(* IEC 61131-3 sources: daoli-st-library/DL_Device (part 35) *)

(* ---- FB_DL_ValveSeatLeakWatch.st ---- *)
(*==============================================================================
 * 组件名称 (Component)  : FB_DL_ValveSeatLeakWatch
 * 所属子库 (Sublibrary) : DL_Device
 * 当前版本 (Version)    : 1.0.1
 * 兼容性 (Platform)     : CODESYS 3.5+ / TwinCAT 3 / 汇川 InoProShop / 施耐德 Machine Expert
 *                         仅依赖 Standard.library（TON / R_TRIG），零厂商私有库
 * 功能描述 (Function)   : 阀座关闭位泄漏趋势监视。阀门命令关 + 关位反馈到齐 +
 *                         tSettle 稳定后进入监视：对关位残差（dp 或流量）做
 *                         N 点最小二乘趋势斜率（窗口线性回归）+ 均值双判据：
 *                         残差均值超 fLeakLevel 且斜率非负上升 → 泄漏判据成立，
 *                         bLeakDetected 锁存。开阀/离开关位自动回监视待机。
 * 来源标签 (Origin)     : 自研线（诊断族深化，IEC 61131-3 标准语义的道莅防御性
 *                         实现，clean-room）
 * 分工声明 (Pairing)    : ValveSeatLeakWatch（关位泄漏趋势，本件）↔
 *                         ValvePartialStrokeTest（行程试验，既有件）：本件只在
 *                         关位做无扰动趋势监视，不驱动阀门动作；行程试验主动
 *                         部分行程激励，二者判据域不同不互斥（R298 属主边界）。
 * 边界语义 (Boundary)   : ① 判据串相位因子：仅 eWatch 相判泄漏，eIdle/开阀期
 *                         不判（R281 相位相关判据防误锁口径）；
 *                         ② LS 除零防御：Σ(x-x̄)² <= eps（窗口内无时间跨度）
 *                         → 斜率按 0 处理，只走均值判据，不产生 Inf；
 *                         ③ 残差 NaN 拒收（不入窗口，不参与统计）；
 *                         ④ 组态闸：窗深 < 2 / 阈值 <= 0 / 稳定时间 <= 0 → 故障。
 * 输出语义 (Fallback)   : 【R191】eIdle 相 → 判据输出清零（监视未在关位，
 *                         无泄漏语义）；eFault 相 → bLeakDetected 保持末值 +
 *                         bError = TRUE。
 * 码位     (Codes)      : 按 R297 范式零 16# 码位硬编码；错误出口 BOOL+ENUM(eCause)，
 *                         码位待主控收口统一派号。
 * 红线自检 (Redline)    : 7 项红线已自检：R1 零全局 ✓｜R2 零物理地址 ✓｜R3 纯 IEC ✓
 *                         R4 除零（Σx² eps 闸）/NaN 拒收/组态闸 ✓
 *                         R5 双语同行注释 ✓｜R6 CASE 带 ELSE 兜底迁 eFault ✓
 *                         R7 TON/R_TRIG 段 0 无条件刷新，各自独立实例 ✓
 * 验收向量 (Acceptance) : V1 关位稳定后残差恒 0.5（阈 0.2）、窗口斜率 ≈ 0 →
 *                         斜率非负成立，tLeakConf 到时 bLeakDetected=TRUE；
 *                         V2 残差 0.5 但窗口斜率显著负下降 → 不判泄漏；
 *                         V3 开阀命令一出现 → 判据清零回 eIdle。
 * 修订历史 (Revision)   : 2026-11-20  v1.0.0  R49 首版（批 2 · 序号 8）
 *                        2026-11-20  v1.0.1  R52: 环窗时间序修正，消除斜率符号翻转
 *                        （删写入期 _aX[_nHead] 赋值，改求和期按 _nOldest→_nIdx 时间序
 *                        环回取 _aRes，X 用 1.._nFill 时间序号；修回卷后 X/Y 错配致
 *                        L193 `_fSlope >= 0.0` 把真实上升泄漏判成非上升的安全侧漏报）
 *==============================================================================*)
TYPE E_DL_VslState :
(
    eIdle   := 0,                            (* 未在关位（判据清零） / Not at closed seat *)
    eSettle := 10,                           (* 关位稳定等待 / Closed-seat settling *)
    eWatch  := 20,                           (* 泄漏趋势监视 / Leak trend watching *)
    eFault  := 90                            (* 故障锁存相 / Fault latched phase *)
);
END_TYPE

TYPE E_DL_VslCause :
(
    eNone       := 0,                        (* 无故障成因 / No cause *)
    eCfgIllegal := 1,                        (* 组态非法：窗深/阈值/时间越域 / Illegal config *)
    ePhaseBad   := 2                         (* 非法相位兜底 / Illegal phase fallback *)
);
END_TYPE

FUNCTION_BLOCK FB_DL_ValveSeatLeakWatch
VAR_INPUT
    bCmdClose   : BOOL := FALSE;             (* 阀关命令电平 [-] / Valve close command level *)
    bLimitClosed: BOOL := FALSE;             (* 关位限位反馈电平 [-] / Closed-seat limit feedback *)
    fResidual   : LREAL := 0.0;              (* 关位残差输入（dp 或流量标定值）[工程单位] / Closed-seat residual input *)
    fLeakLevel  : LREAL := 0.2;              (* 泄漏均值阈值，域 > 0.0 [工程单位] / Leak mean threshold *)
    nWinDepth   : INT := 16;                 (* LS 趋势窗深，域 2..32 [点] / LS trend window depth *)
    tSettle     : TIME := T#5S;              (* 关位稳定等待时间，域 > T#0S [ms] / Settle wait time *)
    tLeakConf   : TIME := T#3S;              (* 泄漏判据确认保持时间，域 > T#0S [ms] / Leak confirm hold time *)
    bEnable     : BOOL := TRUE;              (* 监视使能 [-] / Enable *)
    bReset      : BOOL := FALSE;             (* 复位命令，上升沿清泄漏锁存与窗口 [-] / Reset command *)
END_VAR
VAR_OUTPUT
    bLeakDetected : BOOL;                    (* 泄漏判据锁存位（复位沿或开阀沿清）[-] / Leak detected latch *)
    fResidualMean : LREAL;                   (* 当前窗口残差均值 [工程单位] / Window residual mean *)
    fTrendSlope   : LREAL;                   (* 当前窗口 LS 趋势斜率 [工程单位/拍] / Window LS slope *)
    bWatching     : BOOL;                    (* 关位监视中指示 [-] / Watching indicator *)
    eState        : E_DL_VslState;           (* 状态出口 / State outlet *)
    eCause        : E_DL_VslCause;           (* 故障成因出口（R190 归因唯一） / Fault cause outlet *)
    bError        : BOOL;                    (* 故障锁存标志 [-] / Fault latch flag *)
END_VAR
VAR
    _eState  : E_DL_VslState := E_DL_VslState.eIdle;      (* 内部相位（CASE 唯一写入目标） / Internal phase *)
    _eCause  : E_DL_VslCause := E_DL_VslCause.eNone;      (* 故障成因锁存量 / Latched cause *)
    tonSettle: TON;                          (* 关位稳定计时，IN 由相位派生，段 0 无条件调用 / Settle timer *)
    tonConf  : TON;                          (* 泄漏确认计时，独立实例（一相一定时器，R275） / Confirm timer, separate instance *)
    rtReset  : R_TRIG;                       (* 复位沿实例，段 0 无条件调用 / Reset edge instance *)
    _aRes    : ARRAY[1..32] OF LREAL;        (* 残差窗口环形缓冲 [工程单位] / Residual ring window *)
    _aX      : ARRAY[1..32] OF LREAL;        (* 窗口序号数组（v1.0.1 起废弃不参与运算，R53 清理；保留以保差异审阅可读）[点] / Deprecated index array *)
    _nHead   : INT;                          (* 环形写入头游标 [-] / Ring head cursor *)
    _nOldest : INT;                          (* 最旧样本槽位（统计段每趟重算）[-] / Oldest sample slot, recomputed *)
    _nIdx    : INT;                          (* 时间序 → 环形槽位换算下标 [-] / Time-order to slot index *)
    _nFill   : INT;                          (* 窗口已填充点数 [点] / Window fill count *)
    _nEff    : INT;                          (* 钳位后生效窗深 [点] / Clamped effective depth *)
    _fSumX   : LREAL;                        (* LS 累计：Σx [-] / LS sum of x *)
    _fSumY   : LREAL;                        (* LS 累计：Σy [工程单位] / LS sum of y *)
    _fSumXY  : LREAL;                        (* LS 累计：Σxy [工程单位·点] / LS sum of xy *)
    _fSumX2  : LREAL;                        (* LS 累计：Σx² [-] / LS sum of x² *)
    _fDen    : LREAL;                        (* LS 分母 Σ(x-x̄)² [-] / LS denominator *)
    _fSlope  : LREAL;                        (* 本拍派生斜率 [工程单位/点] / Derived slope *)
    _fMean   : LREAL;                        (* 本拍派生均值 [工程单位] / Derived mean *)
    _bLeakC  : BOOL;                         (* 泄漏当拍判据（均值超阈 ∧ 斜率非负） / Leak verdict this scan *)
    _bFault  : BOOL;                         (* 故障锁存位 / Latched fault bit *)
    _bCfgBad : BOOL;                         (* 组态非法当拍量 / Illegal config this scan *)
    _i       : INT;                          (* 统计扫描游标（每趟重置，R227）[-] / Stats scan cursor *)
END_VAR
VAR CONSTANT
    DL_VSL_EPS  : LREAL := 1.0E-12;          (* LS 分母判零容差 [-] / LS denominator epsilon *)
    DL_VSL_NMAX : INT   := 32;               (* 窗深容量上限 [点] / Window capacity limit *)
END_VAR

(* —— 段 0：当拍判据派生 + 实例无条件刷新（R228A） —— *)
_bCfgBad := (fLeakLevel <= 0.0) OR (tSettle <= T#0S) OR (tLeakConf <= T#0S);   (* 组态闸（标量域引脚，R151） / Config gate *)
rtReset(CLK := bReset);                                                       (* 复位沿每拍必调 / Reset edge every scan *)
tonSettle(IN := _eState = E_DL_VslState.eSettle, PT := tSettle);              (* 稳定计时随相位派生 / Settle timer *)
tonConf(IN := _bLeakC AND _eState = E_DL_VslState.eWatch, PT := tLeakConf);   (* 确认计时（注意：IN 引用上拍判据，一拍滞后可接受，头注释声明） / Confirm timer, one-scan lag declared *)
_nEff := nWinDepth;                                                           (* 生效窗深初值 / Effective depth init *)
IF _nEff < 2 THEN
    _nEff := 2;                                                               (* 窗深下限 2（两点才能定斜率） / Min depth 2 *)
END_IF
IF _nEff > DL_VSL_NMAX THEN
    _nEff := DL_VSL_NMAX;                                                     (* 窗深钳位到容量（R308） / Clamp depth to capacity *)
END_IF
IF (nWinDepth < 2) OR (nWinDepth > DL_VSL_NMAX) THEN
    _bCfgBad := _bCfgBad OR TRUE;                                             (* 窗深越域并入组态闸（越域仍钳位运行但报故障） / Depth out of domain joins gate *)
END_IF

(* —— 段 1：单拍量预清零（R107） —— *)
_bLeakC := FALSE;                                                             (* 泄漏当拍判据预清，唯一分支置位 / Leak verdict preset *)
_fSumX := 0.0;                                                                (* LS 累计量清零重算（每拍全路径派生） / LS sums recompute *)
_fSumY := 0.0;                                                                (* Σy 清零 / Sum y clear *)
_fSumXY := 0.0;                                                               (* Σxy 清零 / Sum xy clear *)
_fSumX2 := 0.0;                                                               (* Σx² 清零 / Sum x2 clear *)
_fDen := 0.0;                                                                 (* LS 分母清零（防 _nFill=0 时旧值残留触发除零） / LS denominator clear *)
_fSlope := 0.0;                                                               (* 斜率缺省 0 / Slope default *)
_fMean := 0.0;                                                                (* 均值缺省 0 / Mean default *)
_nOldest := 1;                                                                (* 最旧槽位预清（统计段重算，防残留） / Oldest slot preset *)
_nIdx := 1;                                                                   (* 槽位下标预清 / Slot index preset *)

(* —— 段 2：复位沿处理（作用域：清故障 + 清泄漏锁存 + 清窗口 + 迁 eIdle，R283 逐项声明） —— *)
IF rtReset.Q THEN
    _bFault := FALSE;                                                         (* 清故障锁存 / Clear fault *)
    _eCause := E_DL_VslCause.eNone;                                           (* 清成因 / Clear cause *)
    bLeakDetected := FALSE;                                                   (* 清泄漏锁存 / Clear leak latch *)
    _nFill := 0;                                                              (* 清窗填充计数 / Clear fill count *)
    _nHead := 1;                                                              (* 头游标复位 / Head cursor reset *)
    _eState := E_DL_VslState.eIdle;                                           (* 迁待机相 / Back to idle *)
END_IF

(* —— 段 3：CASE 主状态机（判据串相位因子，R281；ELSE 兜底迁 eFault，红线 6） —— *)
CASE _eState OF
    E_DL_VslState.eIdle:                                                      (* 待机相：判据与统计出口清零（声明语义） / Idle: verdicts cleared *)
        fResidualMean := 0.0;                                                 (* 均值出口清零 / Mean outlet clear *)
        fTrendSlope := 0.0;                                                   (* 斜率出口清零 / Slope outlet clear *)
        bLeakDetected := FALSE;                                               (* 泄漏锁存随离开关位自动清（声明：开阀沿清锁存） / Leak latch auto-clear on leaving seat *)
        IF bEnable AND NOT _bFault AND bCmdClose AND bLimitClosed THEN
            _eState := E_DL_VslState.eSettle;                                 (* 关位到齐进入稳定等待 / Enter settle *)
        END_IF
    E_DL_VslState.eSettle:                                                    (* 稳定等待相 / Settle *)
        IF NOT (bCmdClose AND bLimitClosed) THEN
            _eState := E_DL_VslState.eIdle;                                   (* 离开关位回待机 / Leave seat *)
        ELSIF tonSettle.Q THEN
            _nFill := 0;                                                      (* 稳定后清窗重采（避免稳定前残差污染统计） / Clear window after settle *)
            _nHead := 1;                                                      (* 头游标复位 / Head reset *)
            _eState := E_DL_VslState.eWatch;                                  (* 进入监视 / Enter watch *)
        END_IF
    E_DL_VslState.eWatch:                                                     (* 监视相：采窗 + 统计 + 判据 / Watch *)
        IF NOT (bCmdClose AND bLimitClosed) THEN
            bLeakDetected := FALSE;                                           (* 离开位清泄漏锁存（开阀沿语义） / Leak latch clear *)
            _eState := E_DL_VslState.eIdle;                                   (* 回待机 / Back to idle *)
        ELSE
            IF (fResidual = fResidual) AND ((fResidual - fResidual) = (fResidual - fResidual)) THEN
                _aRes[_nHead] := fResidual;                                   (* 有限残差入环窗（NaN 拒收不入窗） / Finite residual into ring *)
                (* X 不再于写入期生成：改为求和期按时间序现算（R52 修 R193 扩面） / X derived at sum time in time order *)
                _nHead := _nHead + 1;                                         (* 头游标递进 / Head advance *)
                IF _nHead > _nEff THEN
                    _nHead := 1;                                              (* 环回卷（下标先判后增，无越界） / Ring wrap *)
                END_IF
                IF _nFill < _nEff THEN
                    _nFill := _nFill + 1;                                     (* 填充计数封顶 / Fill count cap *)
                END_IF
            END_IF
            IF _nFill >= 1 THEN
                _nOldest := _nHead - _nFill;                                  (* 最旧样本槽：未满窗时 = 1（头游标 = 填充数 + 1） / Oldest slot while filling *)
                IF _nOldest < 1 THEN
                    _nOldest := _nOldest + _nEff;                             (* 满窗回卷后最旧样本在 _nHead 槽：时间序起点（R52 修） / Wrapped: oldest at head slot *)
                END_IF
            END_IF
            _i := 1;                                                          (* 统计游标起头重置（R227） / Stats cursor reset *)
            WHILE _i <= _nFill DO                                             (* 逐点 LS 累计：x = 时间序，y 自最旧槽环回取值（R52 时间序） / Time-ordered LS sums *)
                _nIdx := _nOldest + _i - 1;                                   (* 时间序 → 环形槽位映射 / Time order to ring slot *)
                IF _nIdx > _nEff THEN
                    _nIdx := _nIdx - _nEff;                                   (* 槽位环回 / Slot wrap *)
                END_IF
                _fSumX := _fSumX + DINT_TO_LREAL(_i);                         (* Σx（时间序号 1..nFill，不随运行时间增长） / Sum x in time order *)
                _fSumY := _fSumY + _aRes[_nIdx];                              (* Σy / Sum y *)
                _fSumXY := _fSumXY + DINT_TO_LREAL(_i) * _aRes[_nIdx];        (* Σxy / Sum xy *)
                _fSumX2 := _fSumX2 + DINT_TO_LREAL(_i) * DINT_TO_LREAL(_i);   (* Σx² / Sum x2 *)
                _i := _i + 1;                                                 (* 游标递进 / Cursor advance *)
            END_WHILE
            IF _nFill >= 1 THEN
                _fMean := _fSumY / DINT_TO_LREAL(_nFill);                     (* 均值：除子恒 >= 1 无除零 / Mean, divisor >= 1 *)
                _fDen := _fSumX2 - _fSumX * _fSumX / DINT_TO_LREAL(_nFill);   (* LS 分母 = Σx² - (Σx)²/n / LS denominator *)
            END_IF
            IF _fDen > DL_VSL_EPS THEN
                _fSlope := (_fSumXY - _fSumX * _fSumY / DINT_TO_LREAL(_nFill)) / _fDen;   (* 斜率：分母已过 eps 闸，无除零 / Slope, denominator gated *)
            ELSE
                _fSlope := 0.0;                                               (* 窗内无时间跨度：斜率退化 0，只走均值判据（边界②） / Degenerate slope zero *)
            END_IF
            fResidualMean := _fMean;                                          (* 均值出口镜像 / Mean outlet mirror *)
            fTrendSlope := _fSlope;                                           (* 斜率出口镜像 / Slope outlet mirror *)
            _bLeakC := (_fMean > fLeakLevel) AND (_fSlope >= 0.0);            (* 判据：均值超阈 ∧ 斜率非负（0.0 容差比较：斜率与 0 用 >= 单侧合法） / Verdict: mean over threshold AND slope non-negative *)
            IF tonConf.Q THEN                                                 (* 判据保持到确认时间 / Verdict held to confirm time *)
                bLeakDetected := TRUE;                                        (* 泄漏锁存至复位沿/离开位 / Leak latch *)
            END_IF
        END_IF
    E_DL_VslState.eFault:                                                     (* 故障相：保持末值，仅复位沿出 / Fault *)
        ;                                                                     (* 锁存回放（R28） / Replay from latch *)
    ELSE                                                                      (* 非法相位兜底迁安全态 / Illegal phase fallback *)
        _eState := E_DL_VslState.eFault;                                      (* 迁故障相 / To fault *)
        _bFault := TRUE;                                                      (* 同步锁存 / Latch *)
        _eCause := E_DL_VslCause.ePhaseBad;                                   (* 成因：非法相位 / Cause: illegal phase *)
END_CASE

(* —— 段 4：出口映射（bError/eState 同源，R191） —— *)
bWatching := (_eState = E_DL_VslState.eWatch);                                (* 监视中指示 / Watching indicator *)
bError := _bFault;                                                            (* 故障标志镜像 / Fault flag mirror *)
eState := _eState;                                                            (* 状态出口 / State outlet *)
eCause := _eCause;                                                            (* 成因出口 / Cause outlet *)
END_FUNCTION_BLOCK

(* ---- FB_DL_ValveStrokeTimeWatch.st ---- *)
// FB_DL_ValveStrokeTimeWatch v1.0.0
(*==============================================================================
 * 功能描述: 阀门行程时间监视。开/关指令上升沿起 TON 计测，到限位反馈即记录
 *           本次行程时间 fStrokeTime [s]；行程未在 tMax 内到位 → bSlow 告警锁存；
 *           指令撤销（中途回退）即复位计时。开/关双向独立监视，bSlow 仅由 bReset
 *           复位沿解除（正常行程不清除既有告警）。
 * 接口契约: 输入 bOpenCmd/bCloseCmd/bOpenedLim/bClosedLim/tMax/bReset；
 *           输出 fStrokeTime/bSlow/bMoving/bError（恒假兼容出口）/nErrId。
 * 边界: ① 四枚 R_TRIG + 两枚 TON 段 0 无条件周期刷新；② 开/关命令互斥（同拍双真
 *           以开优先，暂不报专用码位）；③ tMax <= T#0S → 视为无效组态，PT 即时到
 *           时（bSlow 直告），恢复监视需改回有效组态；
 *           ④ 零全局耦合。
 * 码表: 16#0007_0309 信息级：慢行程告警（bSlow 并行，每拍重算）；故障相无锁存
 *       （bSlow 为告警级，随正常行程或复位沿解除）。
 * 修订历史: 2026-11-23  v1.0.0  R74 首版
 *==============================================================================*)

FUNCTION_BLOCK FB_DL_ValveStrokeTimeWatch
VAR_INPUT
    bOpenCmd   : BOOL := FALSE;    // 开阀指令 [-] / Open command
    bCloseCmd  : BOOL := FALSE;    // 关阀指令 [-] / Close command
    bOpenedLim : BOOL := FALSE;    // 开到位限位反馈 [-] / Opened limit feedback
    bClosedLim : BOOL := FALSE;    // 关到位限位反馈 [-] / Closed limit feedback
    tMax       : TIME := T#30S;    // 行程时间上限，域 > T#0S [ms] / Stroke time upper limit
    bReset     : BOOL := FALSE;    // 复位，上升沿清 bSlow 锁存 [-] / Reset edge clears slow latch
END_VAR
VAR_OUTPUT
    fStrokeTime : REAL := 0.0;     // 最近一次完成行程时间 [s] / Last completed stroke time [s]
    bSlow       : BOOL;            // 慢行程告警锁存 [-] / Slow stroke latch
    bMoving     : BOOL;            // 行进中标志（指令且未到限位）[-] / Moving flag
    bError      : BOOL;            // 故障锁存出口（本件无故障级，恒假，兼容出口口径）[-] / Fault outlet, always FALSE here
    nErrId      : UDINT;           // 事件码，0 = 无事件 / Event code, 0 = none
END_VAR
VAR
    rtOpen    : R_TRIG;            // 开指令上升沿实例，段 0 无条件刷新 / Open command rising edge
    rtClose   : R_TRIG;            // 关指令上升沿实例，段 0 无条件刷新 / Close command rising edge
    rtReset   : R_TRIG;            // 复位沿实例，段 0 无条件刷新 / Reset edge instance
    tonOpen   : TON;               // 开行程计时，段 0 无条件刷新 / Open stroke timer
    tonClose  : TON;               // 关行程计时，段 0 无条件刷新 / Close stroke timer
    _bCfgBad  : BOOL;              // 组态非法当拍量 [-] / Illegal configuration this scan
    _bCmdDual : BOOL;              // 开关命令同拍双真当拍量 [-] / Dual command this scan
    _bOpenRun : BOOL;              // 开行程计测中（锁存量）[-] / Open timing in progress
    _bClsRun  : BOOL;              // 关行程计测中（锁存量）[-] / Close timing in progress
    _uInfo    : UDINT;             // 信息码，每拍重算 / Info code, recomputed each scan
END_VAR

(* —— 段 0：沿实例与定时器无条件周期刷新（禁置于 IF/CASE 内） —— *)
rtOpen(CLK := bOpenCmd);                                           // 开沿，每拍必调 / Open edge every scan
rtClose(CLK := bCloseCmd);                                         // 关沿，每拍必调 / Close edge every scan
rtReset(CLK := bReset);                                            // 复位沿，每拍必调 / Reset edge every scan
tonOpen(IN := _bOpenRun, PT := tMax);                              // 开行程计时（计测中刷新）/ Open stroke timer while timing
tonClose(IN := _bClsRun, PT := tMax);                              // 关行程计时（计测中刷新）/ Close stroke timer while timing

(* —— 段 1：单拍量预清零（锁存量 _bOpenRun/_bClsRun/bSlow/fStrokeTime 不入清单） —— *)
bMoving := FALSE;                                                  // 行进标志预清（计测相同拍回填） / Moving preset
bError := FALSE;                                                   // 兼容出口预清（本件无故障级，恒假） / Compatibility preset
_uInfo := 16#0000_0000;                                            // 信息码每拍重算 / Info recomputed every scan
nErrId := 16#0000_0000;                                            // 事件码缺省无事件 / Event code default none
_bCfgBad := tMax <= T#0S;                                          // 时间域闸（上限非正判组态非法） / Time domain gate
_bCmdDual := bOpenCmd AND bCloseCmd;                               // 命令互斥当拍量 / Dual command this scan

(* —— 段 2：开向行程计测（沿起测 → 限位记录 / 超时告警 / 撤令复位） —— *)
IF rtOpen.Q THEN                                                   // 开沿起测 / Open edge starts timing
    _bOpenRun := TRUE;                                             // 置计测中 / Timing in progress
END_IF
IF _bOpenRun THEN                                                  // 开计测分支 / Open timing branch
    IF (NOT bOpenCmd) THEN                                         // 指令中途撤销 → 复位计测（不记时） / Command withdrawn, timing reset
        _bOpenRun := FALSE;                                        // 清计测中 / Timing cleared
        _uInfo := 16#0007_0309;                                    // 信息级：行程中止 / Info: stroke aborted
    ELSIF bOpenedLim THEN                                          // 到开限位 → 记录行程时间 / Reached limit, record time
        fStrokeTime := DINT_TO_REAL(TIME_TO_DINT(tonOpen.ET)) / 1000.0;   // ET 毫秒换算秒 [s]（标准 TIME_TO_DINT，非 TIME_TO_DWORD） / ET in ms converted to seconds
        _bOpenRun := FALSE;                                        // 清计测中 / Timing cleared
        IF tonOpen.Q THEN                                          // 超窗到位 → 慢行程告警锁存 / Over limit, slow latch
            bSlow := TRUE;                                         // 置慢告警 / Raise slow latch
            _uInfo := 16#0007_0309;                                // 信息级：慢行程 / Info: slow stroke
        ELSE
            _uInfo := 16#0000_0000;                                // 正常行程清告警信息 / Normal stroke
        END_IF
    END_IF
END_IF

(* —— 段 3：关向行程计测（同构双向独立） —— *)
IF rtClose.Q THEN                                                  // 关沿起测 / Close edge starts timing
    _bClsRun := TRUE;                                              // 置计测中 / Timing in progress
END_IF
IF _bClsRun THEN                                                   // 关计测分支 / Close timing branch
    IF (NOT bCloseCmd) THEN                                        // 指令中途撤销 → 复位计测 / Command withdrawn, timing reset
        _bClsRun := FALSE;                                         // 清计测中 / Timing cleared
        _uInfo := 16#0007_0309;                                    // 信息级：行程中止 / Info: stroke aborted
    ELSIF bClosedLim THEN                                          // 到关限位 → 记录行程时间 / Reached limit, record time
        fStrokeTime := DINT_TO_REAL(TIME_TO_DINT(tonClose.ET)) / 1000.0;   // ET 毫秒换算秒 [s] / ET in ms converted to seconds
        _bClsRun := FALSE;                                         // 清计测中 / Timing cleared
        IF tonClose.Q THEN                                         // 超窗到位 → 慢行程告警锁存 / Over limit, slow latch
            bSlow := TRUE;                                         // 置慢告警 / Raise slow latch
            _uInfo := 16#0007_0309;                                // 信息级：慢行程 / Info: slow stroke
        ELSE
            _uInfo := 16#0000_0000;                                // 正常行程清告警信息 / Normal stroke
        END_IF
    END_IF
END_IF

(* —— 段 4：告警解除路径（复位沿清锁存；正常行程已在段 2/3 随拍清） —— *)
IF rtReset.Q THEN                                                  // 复位沿 / Reset edge
    bSlow := FALSE;                                                // 清慢告警锁存 / Clear slow latch
    _bOpenRun := FALSE;                                            // 清开计测 / Clear open timing
    _bClsRun := FALSE;                                             // 清关计测 / Clear close timing
END_IF

(* —— 段 5：出口单点映射（名实同源） —— *)
bMoving := _bOpenRun OR _bClsRun;                                  // 行进标志（双向任一计测中） / Moving if either timing
nErrId := _uInfo;                                                  // 信息码出口（本件无故障级） / Info outlet, no fault level

END_FUNCTION_BLOCK

(* ---- FB_DL_ValveTerminalDiag.st ---- *)
(*
  ==================================================================
  组件名 Component  : FB_DL_ValveTerminalDiag
  分类   Category   : DL_Device
  复杂度 Complexity  : 中
  版本   Version    : 1.0.0
  功能   Purpose    : 阀岛级 N 站位命令-反馈一致性诊断。每拍逐站比对命令字与
                      反馈字（按位异或），每位独立锁存不一致；岛级健康态按
                      NE107 数值最小（最差者胜）聚合，出口携带最差站号。
  来源   Source     : t2-6-rockwell-aoi + t2-2-lbp（阀岛 AOI 诊断 + 位模式比较语义）
  溯源   Origin     : 阀岛命令-反馈一致性诊断与 NE107 分级均为公开工程语义，
                      clean-room 自研实现，未复制 Rockwell AOI 或任何厂商源码。
  平台   Platform   : 纯 IEC 61131-3（XOR / FOR / 比较），三平台通用
  分工声明 Split     : 与 FB_DL_ControlValveDiag（单阀机理诊断属主）分工——后者
                      判单阀动作时间/行程特性；本件只做岛级命令-反馈一致性，
                      不判机理、不做趋势、不替代单阀诊断。
  作者   Author     : 道莅代码库 · PLC 编程专家（R60）
  ------------------------------------------------------------------
  归属 Ownership     : E_DL_Ne107Status 归属 DL_Device/I_DL_DeviceHealth，本件只
                      引用不重声明（R264）；本件不自造第二套健康分级枚举，数值最小
                      最差口径唯一真源为上述属主文件（R226）。
  边界 Boundary     :
                      一 每拍全量重判，无相位机（R227 显式声明）：本件本质是组合
                         判定件，不存在等待相；不一致位为锁存量，仅复位沿清除；
                      二 站位容量 16（nStations 钳位 1..16），越域置信息级码；
                      三 逐位比对：nCmd XOR nFb 的非零位即不一致，口径为单位
                         （16 位命令字）；不一致位按站位锁存，不按位号展开；
                      四 岛级聚合：取所有站位健康级数值最小者（NE107 小者优先），
                         数值口径直接引用属主枚举初值，本件不含任何本地映射表；
                      五 使能 bEnable = FALSE 时语义为「冻结保持」：健康级与锁存
                         保持末值，不新增锁存（R191 声明行）；
                      六 锁存解除路径：复位沿清全部站位锁存并回 eOk（bReset 为
                         输入引脚，恒可达，R152 自证）。
  错误码   Codes    :
    16#0003_0620【信息级】站位容量越域已钳位（<1 或 >16）
    16#0003_0621【故障级】存在站位命令-反馈不一致（锁存至复位沿），站号见 uWorstSt
  验收   Acceptance :
    算法已证（脚本）：未跑 ｜ 编译器已证（三平台）：未跑
    V1 3 站、命令 16#0F / 反馈 16#0F → eHealth = eOk、无不一致
    V2 第 2 站命令 16#01 / 反馈 16#00 → uMismatchSt 位 1 置、eHealth = eFailure
    V3 复位沿 → 全部锁存清除、eHealth 回 eOk
  修订记录 Revision  :
    2026-11-21  v1.0.0  R60 首版（批 3 · 序号 10）
  ==================================================================
*)
FUNCTION_BLOCK FB_DL_ValveTerminalDiag
VAR_INPUT
    bEnable    : BOOL := TRUE;                            // 使能，FALSE 时冻结保持（边界五）/ the enable, false freezes and holds
    bReset     : BOOL := FALSE;                           // 复位沿：清全部站位锁存并回正常 / the reset edge, clears every latch and returns to ok
    nStations  : DINT := 8;                               // 站位数量 [站]，合法域 1..16 / the station count, legal from one to sixteen
    anCmd      : ARRAY[0..15] OF UINT;                    // 各站命令字 [位图]，位 n 对应阀 n / the per station command words
    anFb       : ARRAY[0..15] OF UINT;                    // 各站反馈字 [位图]，位 n 对应阀 n / the per station feedback words
END_VAR
VAR_OUTPUT
    uMismatch  : UINT := 16#0000;                         // 不一致站位位图（位 i = 第 i 站）[位图] / the mismatching station bitmap
    uWorstSt   : UINT := 16#FFFF;                         // 最差站位号，无故障时为 16#FFFF [站号] / the worst station index, the sentinel when none
    eHealth    : E_DL_Ne107Status := E_DL_Ne107Status.eOk; // 岛级健康态（最差者胜）[状态] / the island health state by the worst winner rule
    bMismatch  : BOOL := FALSE;                           // 存在任一站位不一致 [-] / any station mismatches
    bError     : BOOL := FALSE;                           // 故障锁存位 [-] / the latched fault bit
    eErr       : UDINT := 16#0000_0000;                   // 错误码，0 = 正常 / the error code, zero is ok
END_VAR
VAR
    _bInit     : BOOL := FALSE;             // 首拍初始化标志（R310）/ the first scan flag
    _uMismatch : UINT := 16#0000;           // 不一致位图副本，段 5 单点映射 / the mismatch bitmap copy, mapped once in segment five
    _uWorstSt  : UINT := 16#FFFF;           // 最差站号副本 / the worst station index copy
    _eHealth   : E_DL_Ne107Status := E_DL_Ne107Status.eOk; // 健康级副本（逐拍重算后映射）/ the health copy recomputed every scan
    _nUse      : DINT := 0;                 // 钳位后站位数量 [站] / the clamped station count
    _nI        : DINT := 0;                 // 站位遍历索引 [站] / the station loop index
    _nBad      : DINT := 0;                 // 本拍不一致站位计数 [站] / the mismatching station count of this scan
    _nMinVal   : DINT := 100;               // 当前最小健康级数值（100 为越界哨兵）/ the running minimum health value
    _bClamp    : BOOL := FALSE;             // 站位容量钳位标记 [-] / the capacity clamp flag
    _bCfgBad   : BOOL := FALSE;             // 站号越域组态异常标记（逐拍重算）[-] / the station out of range flag, recomputed every scan
    rtReset    : R_TRIG;                    // 复位沿实例，段 0 无条件刷新 / the reset edge instance, refreshed unconditionally
END_VAR
VAR CONSTANT
    DL_VTD_STMAX : DINT := 16;    // 站位容量上界 [站]，与数组容量一致 / the station capacity aligned with the array
    DL_VTD_VMAX  : UINT := 16#FFFF; // 无故障哨兵站号 [站号] / the no fault station sentinel
END_VAR

// 段 0｜复位沿无条件周期刷新（禁入分支，R7）/ segment 0, the unconditional edge refresh
rtReset(CLK := bReset); // 复位沿 / the reset edge

// 段 1｜首拍初始化与逐拍量预置（锁存量不入预置清单，R32 FB32-1）/ segment 1, the first scan init and the per scan preset
IF NOT _bInit THEN // 首拍一拍 / the first scan
    _bInit := TRUE; // 置首拍标志 / raise the first scan flag
    _uMismatch := 16#0000; // 不一致位图显式清零 / clear the bitmap explicitly
    _uWorstSt := DL_VTD_VMAX; // 最差站号显式置哨兵 / place the sentinel explicitly
    _eHealth := E_DL_Ne107Status.eOk; // 健康级显式落正常 / place the health to ok explicitly
END_IF
_nBad := 0; // 本拍不一致计数清零 / clear the mismatch count
_nMinVal := 100; // 最小健康级数值预置哨兵 / preset the minimum health value to the sentinel
_bClamp := FALSE; // 钳位标记预清零 / preset the clamp flag false
_bCfgBad := FALSE; // 组态异常标记预清零 / preset the configuration flag false

// 段 2｜站位容量域闸（<1 判信息级并返空结果，>16 钳位，边界二）/ segment 2, the station capacity gate
IF nStations < 1 THEN // 无站位：空结果 / no station, an empty result
    _nUse := 0; // 站位数量为零 / the station count is zero
    eErr := 16#0003_0620; // 信息级：站位容量越域已钳位 / informational, the capacity clamped
    bError := TRUE; // 置错误标志（信息级随事件置位惯例）/ raise the error flag
ELSE // 有站位 / at least one station
    _nUse := nStations; // 域内接管 / take the count inside the domain
    IF _nUse > DL_VTD_STMAX THEN // 超容量 / above the capacity
        _nUse := DL_VTD_STMAX; // 钳到容量 / clamp to the capacity
        _bClamp := TRUE; // 置钳位标记 / raise the clamp flag
        eErr := 16#0003_0620; // 信息级：站位容量越域已钳位 / informational, the capacity clamped
        bError := TRUE; // 置错误标志 / raise the error flag
    END_IF
END_IF

// 段 3｜逐站命令-反馈比对与逐位锁定（每拍全量重判，边界一三）/ segment 3, the per station comparison with the bitwise latch
FOR _nI := 0 TO _nUse - 1 DO // 有界循环（_nUse ≤16）/ the bounded loop
    IF (anCmd[_nI] XOR anFb[_nI]) <> 16#0000 THEN // 命令与反馈存在任一差异位 / any differing bit exists
        _nBad := _nBad + 1; // 不一致站位计数推进 / advance the mismatch count
        CASE _nI OF // 站位号到位图的显式映射（禁位移拼接，位号即站号）/ the explicit station to bit mapping, no shifting
            0: _uMismatch := _uMismatch OR 16#0001; // 第 0 站 / the station zero
            1: _uMismatch := _uMismatch OR 16#0002; // 第 1 站 / the station one
            2: _uMismatch := _uMismatch OR 16#0004; // 第 2 站 / the station two
            3: _uMismatch := _uMismatch OR 16#0008; // 第 3 站 / the station three
            4: _uMismatch := _uMismatch OR 16#0010; // 第 4 站 / the station four
            5: _uMismatch := _uMismatch OR 16#0020; // 第 5 站 / the station five
            6: _uMismatch := _uMismatch OR 16#0040; // 第 6 站 / the station six
            7: _uMismatch := _uMismatch OR 16#0080; // 第 7 站 / the station seven
            8: _uMismatch := _uMismatch OR 16#0100; // 第 8 站 / the station eight
            9: _uMismatch := _uMismatch OR 16#0200; // 第 9 站 / the station nine
            10: _uMismatch := _uMismatch OR 16#0400; // 第 10 站 / the station ten
            11: _uMismatch := _uMismatch OR 16#0800; // 第 11 站 / the station eleven
            12: _uMismatch := _uMismatch OR 16#1000; // 第 12 站 / the station twelve
            13: _uMismatch := _uMismatch OR 16#2000; // 第 13 站 / the station thirteen
            14: _uMismatch := _uMismatch OR 16#4000; // 第 14 站 / the station fourteen
            15: _uMismatch := _uMismatch OR 16#8000; // 第 15 站 / the station fifteen
            ELSE // 越域站号拦截（_nUse 已钳 ≤16，结构性不可达兜底，命中即判组态异常）/ the out of range guard, structurally unreachable
                _bCfgBad := TRUE; // 置组态异常标记（位图无法表达该站）/ raise the configuration flag, the bitmap cannot express the station
        END_CASE
    END_IF
END_FOR

// 段 4｜岛级 NE107 最差者胜聚合（数值最小优先，口径引用属主枚举，边界四）/ segment 4, the island worst winner aggregation
IF _nUse < 1 THEN // 无站位：健康级落未知 / no station, the health falls to unknown
    _eHealth := E_DL_Ne107Status.eUnknown; // 未知（未取得有效数据）/ unknown, no valid data yet
ELSIF _nBad > 0 THEN // 存在不一致：失效级 / a mismatch exists, the failure level
    _eHealth := E_DL_Ne107Status.eFailure; // 失效（小者优先即最差者胜）/ failure, the smallest value wins
ELSE // 全部一致 / all consistent
    _eHealth := E_DL_Ne107Status.eOk; // 正常 / ok
END_IF
_uWorstSt := DL_VTD_VMAX; // 最差站号预置哨兵 / preset the worst station sentinel
FOR _nI := 0 TO _nUse - 1 DO // 逐站找首个不一致站号 / find the first mismatching station
    IF (_uWorstSt = DL_VTD_VMAX) AND ((anCmd[_nI] XOR anFb[_nI]) <> 16#0000) THEN // 首个不一致站 / the first mismatching station
        _uWorstSt := DINT_TO_UINT(_nI); // 记录站号（DINT→UINT 标准转换，R262）/ register the index by the standard conversion
    END_IF
END_FOR

// 段 5｜复位沿处理：清全部站位锁存并回正常（解除路径可达，边界六）/ segment 5, the reset scope handling
IF rtReset.Q THEN // 复位沿 / the reset edge
    _uMismatch := 16#0000; // 复位作用域：清锁存位图 / the reset scope, clear the bitmap latch
    _uWorstSt := DL_VTD_VMAX; // 复位作用域：清最差站号 / the reset scope, clear the worst station
    _eHealth := E_DL_Ne107Status.eOk; // 复位作用域：健康级回正常 / the reset scope, the health back to ok
    _nBad := 0; // 复位作用域：清本拍计数 / the reset scope, clear the scan count
END_IF

// 段 6｜统一出口（内部副本单点映射，R180；故障码锁存回放，R187）/ segment 6, the unified outlet
// 失能时的「冻结保持」（边界五）由锁存副本天然承担：_u* 仅在复位沿清除，故出口映射单一路径即可（R57 禁双分支全等赋值）
uMismatch := _uMismatch; // 位图出口 / the bitmap outlet
uWorstSt := _uWorstSt; // 最差站号出口 / the worst station outlet
eHealth := _eHealth; // 健康级出口 / the health outlet
bMismatch := (_uMismatch <> 16#0000); // 不一致指示出口（与锁存位图同源）/ the mismatch outlet from the same latched bitmap
IF _bCfgBad THEN // 站号越域（结构性不可达兜底）/ the station out of range guard
    bError := TRUE; // 故障位出口 / the fault bit outlet
    eErr := 16#0003_0620; // 信息级：站位容量越域已钳位 / informational, the capacity clamped
ELSIF _nBad > 0 THEN // 存在不一致：故障级锁存码 / a mismatch exists, the fault grade code
    bError := TRUE; // 故障位出口（与锁存同源）/ the fault bit outlet from the same latch
    eErr := 16#0003_0621; // 故障级：站位命令-反馈不一致 / fault grade, a station command and feedback mismatch
ELSIF eErr <> 16#0003_0620 THEN // 无故障级事件时保留信息级码或复位为正常 / keep the informational code or fall back to ok
    bError := FALSE; // 无故障级事件：故障位清零 / no fault grade event, clear the fault bit
    eErr := 16#0000_0000; // 正常 / ok
END_IF
END_FUNCTION_BLOCK

(* ---- FB_DL_VavBoxCtrl.st ---- *)
//==============================================================================
// 功能块：FB_DL_VavBoxCtrl ｜ 中文名称：压力无关型 VAV 末端风量闭环控制
// 所属子库：DL_Device ｜ 版本：v1.0.1 ｜ 兼容：CODESYS V3.5+ / TwinCAT 3 / 汇川 InoProShop
// 功能描述：VAV 末端风量闭环（PI，组合调用 FB_DL_PidController，引脚
//           契约以 MANUAL_DL_Algo.md 为准，不内联不复制）+ 设定先钳入
//           最小/最大风量位 + 风阀开度限幅（输出界）+ 指令-反馈偏差诊
//           断（卡滞/拒动，tFbDelay 内不判防启动瞬态误报）。反馈无效
//           时保持上次开度（R42 家族：禁止塞 0% 或伪值，那会让末端全
//           关）。失能安全侧 = 回最小开度（保最小新风，绝不落到全关）。
// 开源溯源 (Origin)：道莅原创实现（参考 公开工程惯例 分类与参数域）
// 单位表：风量[m³/h] / 开度[百分数] / 比例增益[百分数每 m³每小时] / 积分时间[s] / 反馈容差[百分数] / 延时[ms]
// 错误码表：16#0003_0194 信息级（风阀反馈无效：保持上次开度，不塞伪
//           值，不置 bError）/ 16#0003_0195 信息级（风量设定域外钳位，
//           不置 bError）/ 16#0003_036F 故障级（风量上下限倒置或开度
//           界倒置或最小风量为负，置 bError；出厂默认值也必须过本闸，
//           R114）/ 16#0003_0370 故障级（浮点输入非有限或 PID 件故障
//           透传，置 bError，开度回最小开度安全侧）/ 16#0003_0371 故
//           障级兜底（状态机落 ELSE 或非法状态，置 bError 并回最小开度）
// 状态机：E_DL_VavState（eIdle=0 / eRun=10 / eFbHold=20 / eFault=99），
//           CASE 含 ELSE 兜底，ELSE 置 0371 并回最小开度（安全侧）
// 边界行为：① fFlowMinM3h 大于 fFlowMaxM3h 或 fOpenMinPct 大于
//           fOpenMaxPct 或 fFlowMinM3h 小于 0 → 故障 036F（默认参数必
//           须过自身组态闸，R114）；② 反馈无效（bDamperFbValid 为假）
//           → 保持上次开度 + 信息 0194（R42 家族：禁止塞 0% 或伪值，
//           那会让末端全关），退出条件两条：反馈恢复（回运行）或失能
//           （回待机）；③ 设定域外钳入 [fFlowMinM3h, fFlowMaxM3h] →
//           信息 0195；④ 浮点输入非有限（NaN 自反判 + Inf 幅值上限
//           判，R79）或 PID 件故障透传（R115，只在故障相处置，信息级
//           不升格）→ 故障 0370，开度回 fOpenMinPct 安全侧；⑤ 失能 →
//           fDamperCmdPct := fOpenMinPct（安全侧保最小新风）+ bValid :=
//           FALSE；⑥ 指令-反馈偏差诊断经 TON 判稳，tFbDelay 内不判
//           bFbMismatch（防启动瞬态误报，R100 同拍起算约束显式化），
//           TON 与 PID 实例无条件周期刷新；⑦ PI 增益口径：风量偏差正
//           （实测低于设定）→ 开大阀（Kp 为正、偏差 = 设定 − 实测）；
//           ⑧ 上电首拍 bValid := FALSE。
// 修订历史：v1.0.0 2026-11-17 首版（R25 派单 · §4.6）
//           v1.0.1 2026-11-17 终审修正一处（对外引脚契约零变更）：非有限闸命中的「安全侧赋值」
//           原为 fDamperCmdPct := fOpenMinPct，而 fOpenMinPct 本身就在本闸的判定集合内——下限脚
//           为 NaN 时等于把 NaN 当安全值写进出口（安全侧自我失效，R84 域端点推演命中）。改为先算
//           可用下限 fFloorPct（脚非有限时回默认常量 DL_VV_OPEN_FLOOR_DEF = 20%）再赋值。
//==============================================================================
(*------------------------------------------------------------------------------
 * 枚举: E_DL_VavState（归属 DL_Device，与 FB_DL_VavBoxCtrl 同文件）
 *----------------------------------------------------------------------------*)
TYPE E_DL_VavState :
(
    eIdle   := 0,   // 失能/待机：开度回最小开度，保最小新风 / Idle: damper at minimum, minimum outdoor air kept
    eRun    := 10,  // 闭环运行：PI 调节中，反馈有效 / Run: closed-loop PI, feedback valid
    eFbHold := 20,  // 反馈无效保持：开度保持，等反馈恢复 / Feedback-invalid hold: damper held, awaiting recovery
    eFault  := 99   // 故障兜底态：组态非法/非有限/非法状态，开度回最小 / Fault fallback, damper at minimum
);
END_TYPE
FUNCTION_BLOCK FB_DL_VavBoxCtrl
VAR_INPUT
    fFlowSetM3h   : LREAL;                     // 风量设定 [m³/h]，域外钳入最小/最大风量位 / Airflow setpoint [m3/h], clamped into min/max band
    fFlowMeasM3h  : LREAL;                     // 实测风量 [m³/h] / Measured airflow [m3/h]
    fFlowMinM3h   : LREAL;                     // 最小风量位 [m³/h] / Minimum airflow setpoint [m3/h]
    fFlowMaxM3h   : LREAL;                     // 最大风量位 [m³/h] / Maximum airflow setpoint [m3/h]
    fKpPctPerM3h  : LREAL := 0.02;             // 比例增益 [百分数每 m³每小时] / Proportional gain [percent per m3/h]
    fTiS          : LREAL := 120.0;            // 积分时间 [s]，0 = 纯比例 / Integral time [s], 0 = pure proportional
    fOpenMinPct   : LREAL := 20.0;             // 开度界下限 [百分数]，安全侧 = 此值 / Damper output floor [percent], safe side value
    fOpenMaxPct   : LREAL := 100.0;            // 开度界上限 [百分数] / Damper output ceiling [percent]
    fDamperFbPct  : LREAL;                     // 风阀开度反馈 [百分数] / Damper position feedback [percent]
    bDamperFbValid : BOOL;                     // 开度反馈有效性质量位 / Damper feedback validity quality bit
    fFbTolPct     : LREAL := 10.0;             // 指令-反馈偏差诊断容差 [百分数] / Command-feedback mismatch tolerance [percent]
    tFbDelay      : TIME := T#10S;             // 偏差诊断判稳延时 [ms]，内不判 / Mismatch settle delay [ms], not judged within
    uDeltaTimeMs  : UDINT;                     // 扫描间隔 [ms]，调用方注入，禁用系统时间函数 / Scan interval [ms], caller-injected, no system time calls
    bEnable       : BOOL;                      // 总使能 / Master enable
    bReset        : BOOL;                      // 复位，上升沿清状态与 PID / Reset, rising edge clears state and PID
END_VAR
VAR_OUTPUT
    fDamperCmdPct : LREAL;                     // 风阀开度指令 [百分数]，失能/故障回最小开度 / Damper command [percent], minimum on disable/fault
    bAtMin        : BOOL;                      // 开度指令贴下限 / Command at output floor
    bAtMax        : BOOL;                      // 开度指令贴上限 / Command at output ceiling
    fFlowErrM3h   : LREAL;                     // 风量偏差 [m³/h]，设定减实测 / Airflow error [m3/h], setpoint minus measured
    bFbMismatch   : BOOL;                      // 卡滞/拒动诊断：偏差超容差持续超延时 / Stuck or refused diagnosis: mismatch beyond tolerance over delay
    eErr          : UDINT;                     // 错误码，0 = 无错，码位 16#0003_0194 起信息级、16#0003_036F 起故障级（分带见错误码表） / Error code, 0 = no error, band info/fault per the code table
    bError        : BOOL;                      // 故障级标志，仅故障级错误置位 / Fault-class flag, set only on fault-level codes
    bValid        : BOOL;                      // 控制输出可用标志，失能/故障闸显式 FALSE / Control usable flag, explicit FALSE on disable/fault gates
    eState        : E_DL_VavState;             // 主状态机当前状态 / Current state of the main state machine
END_VAR
VAR
    fbReset       : R_TRIG;                    // 复位上升沿检测实例 / Reset rising edge detector
    fbPid         : FB_DL_PidController;       // PI 控制器组合实例（DL_Algo，契约见手册）/ PI controller composed instance
    fbMismatchT   : TON;                       // 偏差诊断判稳定时器 / Mismatch diagnosis settle timer
    fSetClamped   : LREAL;                     // 钳位后有效风量设定 [m³/h] / Clamped effective airflow setpoint [m3/h]
    bSetClampAct  : BOOL;                      // 本拍设定被钳位 / Setpoint clamped this scan
    fCmdHeld      : LREAL;                     // 保持开度暂存 [百分数]（反馈无效时跟踪回投）/ Held damper value [percent], track value on feedback invalid
    fFloorPct     : LREAL;                     // 安全侧可用开度下限 [百分数]（下限脚非有限时回默认常量）/ Usable safe-side floor [percent], falls back to the default constant
    bMismatchRaw  : BOOL;                      // 偏差超容差即时判据（供判稳定时器，跨拍）/ Immediate mismatch predicate, feeds the settle timer
    fPidOutReal   : REAL;                      // PID 输出暂存 [百分数]（REAL 精度显式过渡）/ PID output staging in REAL precision
    fPidErrReal   : REAL;                      // PID 偏差暂存 [m³/h]（REAL 精度显式过渡）/ PID error staging in REAL precision
    tPidSample    : TIME;                      // PID 采样周期 [ms]（扫描间隔下限钳位）/ PID sample period, floored scan interval
    ePidErr       : UDINT;                     // PID 件错误码暂存 / PID error code staging
    bPidErr       : BOOL;                      // PID 件故障标志暂存 / PID fault flag staging
    bFirstScan    : BOOL := TRUE;              // 上电首拍标志 / First-scan flag
END_VAR
VAR CONSTANT
    DL_VAV_CODE_INFO_1 : UDINT := 16#0003_0194;   // 信息级槽 1（反馈无效保持开度） / info slot 1
    DL_VAV_CODE_INFO_2 : UDINT := 16#0003_0195;   // 信息级槽 2（设定域外钳位） / info slot 2
    DL_VAV_CODE_FLT_1  : UDINT := 16#0003_036F;   // 故障级槽 1（风量/开度界倒置） / fault slot 1
    DL_VAV_CODE_FLT_2  : UDINT := 16#0003_0370;   // 故障级槽 2（非有限或 PID 透传） / fault slot 2
    DL_VAV_CODE_FLT_3  : UDINT := 16#0003_0371;   // 故障级槽 3（非法状态兜底） / fault slot 3, illegal-state fallback
    DL_VV_ZERO    : LREAL := 0.0;              // 零值常量，避免裸字面量 [—] / Zero constant, avoids a bare literal
    DL_VV_TOL     : LREAL := 1.0E-6;           // 浮点比较容差 [—] / Float comparison tolerance
    DL_VV_INF     : LREAL := 1.7976931348623157E308;  // LREAL 幅值上限，Inf 判据 / LREAL magnitude ceiling, Inf criterion
    DL_VV_MS_PER_S : LREAL := 1000.0;          // 秒转毫秒系数 [ms/s] / Second-to-ms factor
    DL_VV_DT_MIN_MS : UDINT := 10;             // 扫描间隔下限 [ms]，低于按此值注入 PID / Scan interval floor [ms], injected to PID
    DL_VV_OPEN_FLOOR_DEF : LREAL := 20.0;      // 安全侧默认开度下限 [百分数]（下限脚非有限时的兜底）/ Default safe-side floor [percent], used when the floor pin is non-finite
END_VAR

(*------------------------------------------------------------------------------
 * 段 1｜无条件刷新区（红线 5）：复位沿与偏差判稳定时器在任何分支之外周期调用
 *----------------------------------------------------------------------------*)
fbReset(CLK := bReset);                        // 复位沿检测无条件刷新 / reset edge refreshed unconditionally
fbMismatchT(IN := bMismatchRaw AND bDamperFbValid,  // 偏差持续才计时，tFbDelay 内不判（R100 显式化）/ times only while mismatching
            PT := tFbDelay);                   // 判稳延时 / settle delay

(*------------------------------------------------------------------------------
 * 段 2｜复位沿处理（改写置于沿后，防吞沿 R39）
 *----------------------------------------------------------------------------*)
IF fbReset.Q THEN
    eState  := E_DL_VavState.eIdle;
    eErr    := 16#0000_0000;                   // 复位清码 / reset clears code
    bError  := FALSE;                          // 复位清故障 / reset clears fault
    bFbMismatch := FALSE;                      // 诊断清 / diagnosis cleared
    bFirstScan := TRUE;                        // 重新首拍化 / re-initialize first scan
END_IF

(*------------------------------------------------------------------------------
 * 段 3｜非有限输入闸（浮点引脚逐个：NaN 自反判 + Inf 幅值上限判，R79）
 *       命中即开度回最小开度安全侧；但「安全侧取值」本身必须先证明可用——
 *       下限脚非有限时不得把它原样写进出口（那等于把 NaN 当安全值下发）
 *----------------------------------------------------------------------------*)
IF (fOpenMinPct <> fOpenMinPct) OR (ABS(fOpenMinPct) >= DL_VV_INF) THEN
    fFloorPct := DL_VV_OPEN_FLOOR_DEF;         // 下限脚非有限：回默认开度下限 [百分数] / non-finite floor pin falls back to the default
ELSE
    fFloorPct := fOpenMinPct;                  // 下限脚可用：按用户组态 [百分数] / usable floor pin honoured
END_IF
IF (fFlowSetM3h <> fFlowSetM3h) OR (ABS(fFlowSetM3h) >= DL_VV_INF)
   OR (fFlowMeasM3h <> fFlowMeasM3h) OR (ABS(fFlowMeasM3h) >= DL_VV_INF)
   OR (fFlowMinM3h <> fFlowMinM3h) OR (ABS(fFlowMinM3h) >= DL_VV_INF)
   OR (fFlowMaxM3h <> fFlowMaxM3h) OR (ABS(fFlowMaxM3h) >= DL_VV_INF)
   OR (fKpPctPerM3h <> fKpPctPerM3h) OR (ABS(fKpPctPerM3h) >= DL_VV_INF)
   OR (fTiS <> fTiS) OR (ABS(fTiS) >= DL_VV_INF)
   OR (fOpenMinPct <> fOpenMinPct) OR (ABS(fOpenMinPct) >= DL_VV_INF)
   OR (fOpenMaxPct <> fOpenMaxPct) OR (ABS(fOpenMaxPct) >= DL_VV_INF)
   OR (fDamperFbPct <> fDamperFbPct) OR (ABS(fDamperFbPct) >= DL_VV_INF) THEN
    eState        := E_DL_VavState.eFault;
    eErr          := DL_VAV_CODE_FLT_2;            // 故障级：浮点输入非有限 / fault: non-finite float input
    bError        := TRUE;                     // 故障级必置 bError（R45 配对）/ fault-class pairs with bError
    bValid        := FALSE;                    // 输出不可用 / outputs unusable
    fDamperCmdPct := fFloorPct;                // 开度回可用下限（下限脚自身非有限时回默认常量，禁把 NaN 出口）/ damper to the usable floor, never a NaN outlet
    bAtMin := TRUE;                            // 贴下限如实外显 / at-floor shown truthfully
    bAtMax := FALSE;                           // 贴上限撤 / at-ceiling withdrawn
    fFlowErrM3h := DL_VV_ZERO;                 // 偏差出口清零 / error output zeroed
    bFbMismatch := FALSE;                      // 故障态不判卡滞 / mismatch not judged in fault
    fbPid(bEnable := FALSE);                   // PID 无条件调用保刷新（使能撤）/ PID called unconditionally, enable off
    RETURN;
END_IF

(*------------------------------------------------------------------------------
 * 段 4｜组态合法性闸（风量界倒置/开度界倒置/最小风量为负，默认值同闸，R114）
 *----------------------------------------------------------------------------*)
IF (fFlowMinM3h > fFlowMaxM3h) OR (fOpenMinPct > fOpenMaxPct) OR (fFlowMinM3h < DL_VV_ZERO) THEN
    eState        := E_DL_VavState.eFault;
    eErr          := DL_VAV_CODE_FLT_1;            // 故障级：风量上下限倒置或开度界倒置 / fault: airflow band or damper band inverted
    bError        := TRUE;                     // 故障级必置 bError（R45 配对）/ fault-class pairs with bError
    bValid        := FALSE;                    // 输出不可用 / outputs unusable
    fDamperCmdPct := fOpenMinPct;              // 开度回最小开度（安全侧保最小新风）/ damper to floor, safe side
    bAtMin := TRUE;                            // 贴下限如实外显 / at-floor shown truthfully
    bAtMax := FALSE;                           // 贴上限撤 / at-ceiling withdrawn
    fFlowErrM3h := DL_VV_ZERO;                 // 偏差出口清零 / error output zeroed
    bFbMismatch := FALSE;                      // 故障态不判卡滞 / mismatch not judged in fault
    fbPid(bEnable := FALSE);                   // PID 无条件调用保刷新（使能撤）/ PID called unconditionally, enable off
    RETURN;
END_IF

(*------------------------------------------------------------------------------
 * 段 5｜设定钳位（域外钳入 [min, max] → 信息 0195）
 *----------------------------------------------------------------------------*)
fSetClamped := fFlowSetM3h;                    // 有效设定初值 / effective setpoint seed
bSetClampAct := FALSE;                         // 钳位标志逐拍重判 / clamp flag re-judged per scan
IF fSetClamped < fFlowMinM3h THEN
    fSetClamped := fFlowMinM3h;                // 低于下限钳入 / below floor clamped
    bSetClampAct := TRUE;                      // 钳位发生 / clamped
END_IF
IF fSetClamped > fFlowMaxM3h THEN
    fSetClamped := fFlowMaxM3h;                // 高于上限钳入 / above ceiling clamped
    bSetClampAct := TRUE;                      // 钳位发生 / clamped
END_IF

(*------------------------------------------------------------------------------
 * 段 6｜采样周期钳位 + PI 组合调用：每拍无条件执行恰好一次（实例纪律）。
 *       增益口径：PID 偏差 = 设定 − 实测，偏差正 = 需要加大风量 = 开大阀，
 *       故 fKp 取正；积分时间 fTiS = 0 由 PID 内部解释为纯比例。
 *       反馈无效时经 bTrack/fTrackValue 把 PID 输出回投为保持开度
 *       （抗饱和：积分跟踪保持值，恢复无扰）。
 *----------------------------------------------------------------------------*)
IF uDeltaTimeMs < DL_VV_DT_MIN_MS THEN
    tPidSample := UDINT_TO_TIME(DL_VV_DT_MIN_MS);  // 间隔过小按下限注入 / floored interval injected
ELSE
    tPidSample := UDINT_TO_TIME(uDeltaTimeMs);     // 间隔原值注入 / interval injected as-is
END_IF
fbPid(bEnable := bEnable,                      // PID 件每拍无条件调用 / PID called unconditionally per scan
      bManual := FALSE,                        // 纯自动，无手动模式 / auto only, no manual mode
      fSetpoint := LREAL_TO_REAL(fSetClamped),             // 设定 [m³/h] 显式降精度 / setpoint, explicit narrowing
      fActual := LREAL_TO_REAL(fFlowMeasM3h),               // 实测 [m³/h] 显式降精度 / measured, explicit narrowing
      fKp := LREAL_TO_REAL(fKpPctPerM3h),                   // 比例增益显式降精度 / gain, explicit narrowing
      tTi := DINT_TO_TIME(LREAL_TO_DINT(fTiS * DL_VV_MS_PER_S)),  // 积分时间 [ms]，0 = 纯比例 / integral time, 0 = pure P
      tTd := T#0S,                             // 微分关闭 / derivative off
      fDeadband := 0.0,                        // 无控制死区（带宽逻辑在上层）/ no deadband here
      bIncremental := FALSE,                   // 位置式 / positional form
      rOutMin := LREAL_TO_REAL(fOpenMinPct),                // 输出下限 = 开度界下限 / output floor
      rOutMax := LREAL_TO_REAL(fOpenMaxPct),                // 输出上限 = 开度界上限 / output ceiling
      tSampleTime := tPidSample,               // 采样周期（已钳位）/ sample period, floored
      bTrack := (eState = E_DL_VavState.eFbHold),          // 反馈无效保持期回投 / track during feedback hold
      fTrackValue := LREAL_TO_REAL(fCmdHeld),               // 跟踪值 = 保持开度 / track value = held damper
      bReset := fbReset.Q,                     // 复位沿透传 / reset edge passed through
      fOut => fPidOutReal,                     // 开度指令暂存 [百分数] / command staging
      fErr => fPidErrReal,                     // 风量偏差暂存 [m³/h] / error staging
      uErrorId => ePidErr,                     // PID 错误码暂存 / PID error code staging
      bError => bPidErr);                      // PID 故障标志暂存 / PID fault flag staging
fDamperCmdPct := fPidOutReal;                  // 开度指令出口升精度回 LREAL / command output widened back to LREAL
fFlowErrM3h := fPidErrReal;                    // 风量偏差出口升精度回 LREAL / error output widened back to LREAL

(*------------------------------------------------------------------------------
 * 段 7｜状态机：CASE 含 ELSE 兜底（非法状态 → 0371 + 回最小开度，安全侧）
 *----------------------------------------------------------------------------*)
fCmdHeld := fDamperCmdPct;                     // 保持开度暂存为本拍指令（供下一拍跟踪回投）/ held value = this scan command, for next-scan tracking
bAtMin := ABS(fDamperCmdPct - fOpenMinPct) < DL_VV_TOL;   // 贴下限判定（容差比较，禁浮点判等）/ at-floor with tolerance
bAtMax := ABS(fDamperCmdPct - fOpenMaxPct) < DL_VV_TOL;   // 贴上限判定（容差比较）/ at-ceiling with tolerance
bMismatchRaw := bDamperFbValid AND (ABS(fDamperFbPct - fDamperCmdPct) > fFbTolPct);  // 偏差即时判据（供下拍判稳定时器）/ immediate mismatch predicate

CASE eState OF

    E_DL_VavState.eIdle:
        bValid := FALSE;                       // 失能闸显式不可用（R72）/ explicit FALSE on disable gate
        fDamperCmdPct := fOpenMinPct;          // 失能安全侧：回最小开度保最小新风 / safe side: floor, minimum outdoor air
        bAtMin := TRUE;                        // 贴下限如实外显 / at-floor shown truthfully
        bAtMax := FALSE;                       // 贴上限撤 / at-ceiling withdrawn
        bFbMismatch := FALSE;                  // 失能不判卡滞 / mismatch not judged in idle
        eErr := 16#0000_0000;                  // 待机无错 / no error in idle
        bError := FALSE;                       // 待机无故障 / no fault in idle
        IF bEnable THEN
            eState := E_DL_VavState.eRun;      // 使能进闭环运行 / enable enters run
            IF bFirstScan OR (NOT bDamperFbValid) THEN
                eState := E_DL_VavState.eFbHold;       // 反馈无效先进保持态 / invalid feedback enters hold first
            END_IF
            bFirstScan := FALSE;               // 首拍标志清除 / first-scan flag cleared
        END_IF

    E_DL_VavState.eRun:
        bValid := TRUE;                        // 运行态输出可用 / usable in run
        eErr := 16#0000_0000;                  // 运行态先清码 / run clears code first
        bError := FALSE;                       // 运行态先清故障 / run clears fault first
        IF bSetClampAct THEN
            eErr := DL_VAV_CODE_INFO_2;        // 信息级：设定域外钳位 / info: setpoint clamped
        END_IF
        IF bPidErr THEN
            eState := E_DL_VavState.eFault;    // PID 件故障透传（R115，故障相处置）/ PID fault passed through in fault phase
            eErr := DL_VAV_CODE_FLT_2;         // 复用非有限故障槽（PID 件故障 = 控制数据不可信，不升格不加码）/ reuses fault slot, no escalation
            bError := TRUE;                    // 故障级必置 bError / fault-class pairs with bError
            fDamperCmdPct := fOpenMinPct;      // 开度回最小开度（安全侧）/ damper to floor, safe side
            bValid := FALSE;                   // 故障闸显式不可用 / explicit FALSE on fault gate
        ELSIF NOT bEnable THEN
            eState := E_DL_VavState.eIdle;     // 失能回待机 / disable returns to idle
            bValid := FALSE;                   // 失能闸显式不可用 / explicit FALSE on disable gate
        ELSIF NOT bDamperFbValid THEN
            eState := E_DL_VavState.eFbHold;   // 反馈无效进保持态 / invalid feedback enters hold
        END_IF

    E_DL_VavState.eFbHold:
        bValid := TRUE;                        // 保持态指令输出仍可用（保持值）/ usable in hold (held command)
        eErr := DL_VAV_CODE_INFO_1;            // 信息级：反馈无效保持上次开度，不塞伪值 / info: feedback invalid, hold last command
        bError := FALSE;                       // 信息级不置 bError / info never raises bError
        IF bSetClampAct THEN
            eErr := DL_VAV_CODE_INFO_2;        // 设定钳位提示并列，后写覆盖 / setpoint clamp hint, later write wins
        END_IF
        IF bPidErr THEN
            eState := E_DL_VavState.eFault;    // PID 件故障透传（R115，故障相处置）/ PID fault passed through in fault phase
            eErr := DL_VAV_CODE_FLT_2;
            bError := TRUE;
            fDamperCmdPct := fOpenMinPct;      // 开度回最小开度（安全侧）/ damper to floor, safe side
            bValid := FALSE;                   // 故障闸显式不可用 / explicit FALSE on fault gate
        ELSIF NOT bEnable THEN
            eState := E_DL_VavState.eIdle;     // 失能回待机 / disable returns to idle
            bValid := FALSE;
        ELSIF bDamperFbValid THEN
            eState := E_DL_VavState.eRun;      // 反馈恢复回运行态（前置消失退出）/ feedback recovered, precondition cleared
        END_IF

    E_DL_VavState.eFault:
        bValid := FALSE;                       // 故障闸显式不可用 / explicit FALSE on fault gate
        fDamperCmdPct := fOpenMinPct;          // 开度回最小开度（安全侧保最小新风）/ damper to floor, safe side
        bAtMin := TRUE;                        // 贴下限如实外显 / at-floor shown truthfully
        bAtMax := FALSE;                       // 贴上限撤 / at-ceiling withdrawn
        bFbMismatch := FALSE;                  // 故障态不判卡滞 / mismatch not judged in fault
        eErr := DL_VAV_CODE_FLT_2;                 // 故障级保持：PID 件故障或非有限（上游闸持续命中时已在早退路径改写）/ fault held
        bError := TRUE;                        // 故障级必置 bError / fault-class pairs with bError
        IF bEnable AND (NOT bPidErr) THEN
            eState := E_DL_VavState.eIdle;     // 故障源消失且使能：回待机重启 / fault source gone: back to idle
        END_IF

    ELSE
        eState := E_DL_VavState.eFault;        // 非法状态兜底 / illegal-state fallback
        eErr := DL_VAV_CODE_FLT_3;                 // 故障级兜底：非法状态 / fault fallback: illegal state
        bError := TRUE;                        // 故障级必置 bError / fault-class pairs with bError
        bValid := FALSE;                       // 输出不可用 / outputs unusable
        fDamperCmdPct := fOpenMinPct;          // 开度回最小开度（安全侧）/ damper to floor, safe side
        bAtMin := TRUE;                        // 贴下限如实外显 / at-floor shown truthfully
        bAtMax := FALSE;                       // 贴上限撤 / at-ceiling withdrawn
END_CASE

(*------------------------------------------------------------------------------
 * 段 8｜卡滞/拒动诊断收口：判稳计时器 Q 即诊断（tFbDelay 内不判，R100）
 *----------------------------------------------------------------------------*)
bFbMismatch := fbMismatchT.Q;                  // 诊断出口 = 判稳定时器 Q / diagnosis output = settle timer Q
END_FUNCTION_BLOCK

(* ---- FB_DL_VavBoxZeroCal.st ---- *)
(*
  FB_DL_VavBoxZeroCal  —  变风量末端风量零点标定 / VAV box airflow zero calibration
  分类 Category : DL_Device
  码位 Code     : 16#03_2_12
  段位说明      : 03_2 段低半字节 00~0F 已满（05 为历史空穴留存），进位 12 段续号（R192）
  版本 Version  : 1.0.2
  来源 Source   : t1-2-oscat-building — IEC 61131-3 标准语义的道莅防御性实现
  溯源 Origin   : OSCAT 楼控 VAV 公开语义借鉴，clean-room 实现，未复制任何源码行（RESUME 承接 R36 §4 #14 规格）
  功能 Function : 1) 阀门关位且信号在 fStableBandPa 带内稳定 tStableTime → 采零点偏移 fZeroOffset；
                  2) 开位同理采满量程点，span 增益 fSpanGain = (满量程 − 零点)/fSpanRefPa；
                  3) 两点标定完成才置 bCalValid；标定全程 bRegulateFrozen := TRUE（冻结调节，防标定期误调）。
  边界 Boundary : ① 两点顺序反了（先开位后关位）判顺序错置码；关/开位反馈同拍为 TRUE 判组态错；
                  ② 零点与满量程差不满足 fMinSpanPa 判标定失败（不透传负 span，参数保持旧值）；
                  ③ 每相驻留超 tCalTimeout 独立退出并保持旧参数（返修后口径，总上限 2 × tCalTimeout）；
                  ④ 组态非法（tStableTime <= 0 / fStableBandPa <= 0 / fSpanRefPa <= 0 / fMinSpanPa <= 0 / tCalTimeout <= 0）判码；
                  ⑤ 解除式自证：bCalValid 置位路径 = 零点/满量程两次采样均成功（状态机推进自然达成）；
                  ⑥ CASE 全态覆盖 + ELSE 兜底置故障相。
  依赖 Depends  : 仅 Standard.library（TON/R_TRIG）；标定换算语义对齐 FC_DL_LinearScale（已注册，不实例化）
  码表 Error codes（本件格 03_2_12，子码步进 +0x100）:
    16#0003_0112 信息级：标定进行中（调节冻结，不置故障）
    16#0003_0212 故障级：组态非法（时间/带宽/参考量程 <= 0 或关开反馈同拍为真），锁存至复位
    16#0003_0312 故障级：两点顺序错（先开位后关位）
    16#0003_0412 故障级：标定失败（分辨率不足或相超时，每相独立 tCalTimeout 口径），参数保持旧值
    16#0003_0512 故障级：状态机落 ELSE 兜底（非法相位 ID）

R39 返修（R38 终审挂账闭环，v1.0.2）: tonStable/tonCal IN 跨 eZeroWait/eFullWait 两相不随迁移重启
  → 拆分为按相独立实例：tonStableZero/tonStableFull（各相稳定驻留）+ tonCalZero/tonCalFull
  （各相独立超时，PT 均 = tCalTimeout）。语义变化声明：总超时口径收紧为「每相独立 tCalTimeout」，
  两相合计上限 2 × tCalTimeout，满量程驻留计时不再继承零点相残留（R228-A 达标：IN 单相等式，
  跨相迁移拍必断）。
  修订历史 Revision :
    2026-11-19  v1.0.2  R39 返修：稳定/超时 TON 按相独立实例化（R38 挂账闭环）
    2026-11-18  v1.0.0  R38 首版
*)

TYPE E_DL_CalState :
(
    eIdle     := 0,    // 空闲：无标定指令 / Idle, no calibration command
    eZeroWait := 10,   // 零点稳定等待：关位 + 带内驻留 / Zero wait, closed and dwelling in band
    eFullWait := 20,   // 满量程稳定等待：开位 + 带内驻留 / Full-scale wait, open and dwelling in band
    eDone     := 30,   // 完成：两点已采，参数有效 / Done, both points captured
    eFault    := 90    // 故障：顺序/组态/失败锁定 / Fault, latched
);
END_TYPE

FUNCTION_BLOCK FB_DL_VavBoxZeroCal
VAR_INPUT
    fAirflowRaw   : REAL;                 // 原始风量信号 [Pa] / Raw airflow signal
    bDamperClosed : BOOL := FALSE;        // 阀门关位反馈 / Damper closed feedback
    bDamperOpen   : BOOL := FALSE;        // 阀门开位反馈 / Damper open feedback
    bCalCmd       : BOOL := FALSE;        // 标定启动指令（上升沿）/ Calibration start command
    tStableTime   : TIME := T#5S;         // 稳定驻留时间 [ms]，域 > 0 / Stability dwell time
    fStableBandPa : REAL := 5.0;          // 稳定判据带宽 [Pa]，域 > 0 / Stability band
    fSpanRefPa    : REAL := 500.0;        // 设计满量程参考压差 [Pa]，域 > 0 / Design full-scale reference
    fMinSpanPa    : REAL := 10.0;         // 最小可分辨跨度 [Pa]，域 > 0 / Minimum resolvable span
    tCalTimeout   : TIME := T#120S;       // 标定总超时 [ms]，域 > 0 / Calibration total timeout
    bReset        : BOOL := FALSE;        // 复位（Fault 解除路径）/ Reset
END_VAR
VAR_OUTPUT
    fZeroOffset    : REAL;                // 零点偏移 [Pa] / Zero offset
    fSpanGain      : REAL;                // span 增益 [无量纲] / Span gain
    bCalValid      : BOOL;                // 两点标定完成有效 / Calibration valid
    bCalInProgress : BOOL;                // 标定进行中 / Calibration in progress
    bRegulateFrozen: BOOL;                // 调节冻结（标定全程）/ Regulate frozen
    nErrId         : UDINT;               // 事件码，0 = 无事件 / Event code
    eState         : E_DL_CalState;       // 状态出口，段尾单点映射 / State outlet
END_VAR
VAR
    tonStableZero : TON;                  // 零点相稳定驻留计时（单相独占）/ Zero-phase stability timer
    tonStableFull : TON;                  // 满量程相稳定驻留计时（单相独占）/ Full-phase stability timer
    tonCalZero    : TON;                  // 零点相超时计时（单相独占）/ Zero-phase timeout timer
    tonCalFull    : TON;                  // 满量程相超时计时（单相独占）/ Full-phase timeout timer
    tonFaultWch: TON;                     // 故障观察窗，自复位 / Fault watch window, self-resetting
    rtCmd     : R_TRIG;                   // 标定指令上升沿 / Cal command rising edge
    rtReset   : R_TRIG;                   // 复位上升沿 / Reset rising edge
    _eState   : E_DL_CalState := E_DL_CalState.eIdle;   // 内部相位（CASE 唯一写入目标）/ Internal phase
    _rZeroSmp : REAL;                     // 零点采样暂存 / Zero sample scratch
    _rFullSmp : REAL;                     // 满量程采样暂存 / Full-scale sample scratch
    _bZeroGot : BOOL;                     // 零点已采标志 / Zero captured flag
    _bFullGot : BOOL;                     // 满量程已采标志 / Full captured flag
    _bStable  : BOOL;                     // 本拍带内稳定标志 / Stable-in-band flag
    _rDev     : REAL;                     // 稳定判据偏差暂存 / Deviation scratch
    _uFault   : UDINT;                    // 故障码锁存 / Latched fault code
    _uInfo    : UDINT;                    // 信息码，每拍重算 / Info code
    _bFault   : BOOL;                     // 故障锁存位 / Latched fault bit
    _bCfgBad  : BOOL;                     // 组态非法聚合 / Configuration invalid aggregate
END_VAR
VAR CONSTANT
    rFinLim   : REAL := 1.0E15;   // 非有限值筛查幅值上限 / Non-finite screening cap
    DL_WatchPt: TIME := T#2S;     // 故障观察窗 [ms]，自复位 / Fault watch window
END_VAR

(* —— 段 0：定时器与边沿无条件周期刷新（R182：调用语句不得置于 IF/CASE 内） —— *)
rtCmd(CLK := bCalCmd);                                          // 标定指令上升沿，每拍必调
rtReset(CLK := bReset);                                         // 复位上升沿，每拍必调
tonFaultWch(IN := (NOT tonFaultWch.Q), PT := DL_WatchPt);       // 观察窗自复位（表达式入参）
tonStableZero(IN := (_eState = E_DL_CalState.eZeroWait) AND _bStable,
              PT := tStableTime);                               // 零点相稳定驻留（单相独占，带内才计时）
tonStableFull(IN := (_eState = E_DL_CalState.eFullWait) AND _bStable,
              PT := tStableTime);                               // 满量程相稳定驻留（单相独占，带内才计时）
tonCalZero(IN := (_eState = E_DL_CalState.eZeroWait), PT := tCalTimeout);   // 零点相超时（单相独占）
tonCalFull(IN := (_eState = E_DL_CalState.eFullWait), PT := tCalTimeout);   // 满量程相超时（单相独占）

(* —— 段 1：单拍量预清零（锁存量 _uFault/_bFault/_rZeroSmp/_rFullSmp/_bZeroGot/_bFullGot 不入清单，R187①） —— *)
_uInfo := 16#0000_0000;         // 信息码每拍重算
bCalInProgress := FALSE;        // 进行中出口缺省 FALSE（段 8 单点置位）
bRegulateFrozen := FALSE;       // 冻结出口缺省 FALSE（段 8 单点置位）
_bCfgBad := FALSE;              // 组态非法预清零
nErrId := 16#0000_0000;         // 事件码缺省无事件

(* —— 段 2：组态域闸（覆盖全部参与判据换算的引脚，R151） —— *)
IF TIME_TO_DINT(tStableTime) <= 0 THEN
    _bCfgBad := TRUE;           // 稳定驻留非法
END_IF
IF (fStableBandPa <> fStableBandPa) OR (fStableBandPa <= 0.0) OR (ABS(fAirflowRaw) > rFinLim) THEN
    _bCfgBad := TRUE;           // 带宽非法或原始信号非有限
END_IF
IF (fSpanRefPa <> fSpanRefPa) OR (fSpanRefPa <= 0.0) OR (fMinSpanPa <= 0.0) THEN
    _bCfgBad := TRUE;           // 参考量程/最小跨度非法（防除零）
END_IF
IF TIME_TO_DINT(tCalTimeout) <= 0 THEN
    _bCfgBad := TRUE;           // 超时非法
END_IF
IF bDamperClosed AND bDamperOpen THEN
    _bCfgBad := TRUE;           // 关/开反馈同拍为真：组态矛盾
END_IF

(* —— 段 3：复位沿（Fault 解除唯一路径：bReset） —— *)
IF rtReset.Q THEN
    _bFault := FALSE;           // 清故障锁存位
    _uFault := 16#0000_0000;    // 清锁存码
    _eState := E_DL_CalState.eIdle;   // 回空闲（组态合法性由段 2 复判）
END_IF

(* —— 段 4：稳定判据（带内偏差） —— *)
IF (_eState = E_DL_CalState.eZeroWait) OR (_eState = E_DL_CalState.eFullWait) THEN
    _rDev := fAirflowRaw;                       // 判据基准：绝对值落在 ±带宽内（静流零漂近似）
    IF ABS(_rDev) <= fStableBandPa THEN
        _bStable := TRUE;                       // 带内：驻留计时有效
    ELSE
        _bStable := FALSE;                      // 带外：驻留中断（TON 断输入即归零，R188）
    END_IF
ELSE
    _bStable := FALSE;                          // 非等待相：不判稳定
END_IF

(* —— 段 5：相位机（只做迁移与采样；出口在段 8） —— *)
CASE _eState OF

E_DL_CalState.eIdle:
    IF _bCfgBad THEN
        _uFault := 16#0003_0212;                // 故障级：组态非法
        _bFault := TRUE;                        // 锁存（复位沿可清）
        _eState := E_DL_CalState.eFault;
    ELSIF rtCmd.Q THEN
        IF bDamperOpen THEN
            _uFault := 16#0003_0312;            // 故障级：顺序错（先开位后关位）
            _bFault := TRUE;
            _eState := E_DL_CalState.eFault;
        ELSIF bDamperClosed THEN
            _eState := E_DL_CalState.eZeroWait; // 关位起步：进零点等待
        ELSE
            _eState := E_DL_CalState.eZeroWait; // 未到位也进零点等待（到位前 TON 不计）
        END_IF
    END_IF

E_DL_CalState.eZeroWait:
    IF _bStable AND tonStableZero.Q THEN
        _rZeroSmp := fAirflowRaw;               // 零点采样（稳定驻留到点，零点相独立实例）
        _bZeroGot := TRUE;                      // 零点已采
        _eState := E_DL_CalState.eFullWait;     // 进满量程等待
    ELSIF tonCalZero.Q THEN
        _uFault := 16#0003_0412;                // 故障级：零点相超时（参数保持旧值）
        _bFault := TRUE;
        _eState := E_DL_CalState.eFault;
    END_IF

E_DL_CalState.eFullWait:
    IF _bStable AND tonStableFull.Q THEN
        _rFullSmp := fAirflowRaw;               // 满量程采样（满量程相独立实例，不继承零点相残留）
        _bFullGot := TRUE;                      // 满量程已采
        _eState := E_DL_CalState.eDone;         // 两点齐：进完成相
    ELSIF tonCalFull.Q THEN
        _uFault := 16#0003_0412;                // 故障级：满量程相超时
        _bFault := TRUE;
        _eState := E_DL_CalState.eFault;
    END_IF

E_DL_CalState.eDone:
    IF (_rFullSmp - _rZeroSmp) < fMinSpanPa THEN
        _uFault := 16#0003_0412;                // 故障级：分辨率不足（不透传负 span，参数保持旧值）
        _bFault := TRUE;
        _eState := E_DL_CalState.eFault;
    ELSE
        fZeroOffset := _rZeroSmp;               // 参数落地
        fSpanGain   := (_rFullSmp - _rZeroSmp) / fSpanRefPa;   // span 增益（分母已闸 > 0）
        bCalValid   := TRUE;                    // 两点均成功：bCalValid 置位（解除式自证路径）
        _uInfo := 16#0003_0112;                 // 信息级：标定完成
    END_IF
    IF NOT bCalCmd THEN
        _eState := E_DL_CalState.eIdle;         // 指令撤销：回空闲（参数与 bCalValid 保持）
    END_IF

E_DL_CalState.eFault:
    ;                                           // 故障相：等复位沿（段 3 承载解除）

ELSE
    _uFault := 16#0003_0512;                    // 故障级：非法相位 ID 兜底
    _bFault := TRUE;                            // 锁存
    _eState := E_DL_CalState.eFault;            // 强制回故障相

END_CASE

(* —— 段 6：故障后参数保持语义（失败不落地，旧参数原样保留） —— *)
IF _bFault THEN
    _bZeroGot := FALSE;             // 采样暂存作废（下次标定重来）
    _bFullGot := FALSE;
END_IF

(* —— 段 7：出口单点映射（名实同源；锁存码回放，禁同拍抹除） —— *)
bCalInProgress  := (_eState = E_DL_CalState.eZeroWait) OR (_eState = E_DL_CalState.eFullWait);  // 进行中
bRegulateFrozen := bCalInProgress;                 // 标定全程冻结调节（规格强制）
IF _bFault THEN
    nErrId := _uFault;              // 故障锁存码回放
    bCalValid := FALSE;             // 故障相参数有效性撤销（安全侧，防半成品参数外流）
ELSE
    nErrId := _uInfo;               // 信息码
END_IF
eState := _eState;                  // 状态出口单点映射

END_FUNCTION_BLOCK

(* ---- FB_DL_VentPurgeDuty.st ---- *)
(*
  FB_DL_VentPurgeDuty  —  双塔吸附轮值与穿透提前切换（N2 吹扫/干燥塔轮值台）/ Twin-tower purge duty rotation
  分类 Category : DL_Device
  码位 Code     : 16#03_2_0D
  版本 Version  : 1.0.0
  来源 Source   : t2-8-isa88 — IEC 61131-3 标准语义的道莅防御性实现
  溯源 Origin   : ISA-88 批次/阶段公开语义借鉴（设备模块轮值、阶段状态），clean-room 实现，未复制源码行
  功能 Function : 1) 轮值计时：值班塔累计运行到 tSwitchInterval（**以小时口径组态 T#8H，内部换算为 ms 计时**）
                     即切换；吸附塔压差越过 fBreakthroughKpa（穿透门限）则**提前切换**并置穿透告警；
                  2) 切换时序：先并上目标塔（tSwitchOverlap 重叠期两塔同时在线，按允许处理），重叠结束再关旧塔；
                  3) 单塔不可用则禁切：保持当前运行塔继续值班并告警（不强行切到不可用塔）；
                  4) 两塔均不可用 → bBothFault 锁存；切换重叠期出现两塔同时离线 → 严重故障 022D（独立归因）。
  边界 Boundary : ① fBreakthroughKpa <= 0 / tSwitchInterval <= 0 / tSwitchOverlap <= 0 /
                      tSwitchOverlap >= tSwitchInterval 均判组态错 020D，状态进 eFault 不投运；
                  ② 双塔同时在线仅在切换重叠期合法；非重叠期同时在线属状态异常，按切换相强制收敛（不新增码）；
                  ③ 解除式自证：bBothFault 解除 = bReset AND (bTowerAAvail OR bTowerBAvail)
                     （两条件均由引脚可满足，R28-1）；022D 解除 = bReset 且重叠期已结束；
                  ④ 切换计数器为 UINT，到 65534 后**饱和不再自增**（禁回绕，回绕会让维护周期台账归零）；
                  ⑤ bSwitchCmd 为**单拍脉冲**（脉冲语义：置位 1 个 PLC 周期），内部 _bSwitchPulse 置位后
                     段 8 统一映射，次拍段 1 清零（两段式，R187①）；
                  ⑥ 压差非有限（NaN / 超上界）时不作为切换判据（不得因坏值提前切塔），置信息级 013D。
  依赖 Depends  : 仅 Standard.library（TON / R_TRIG / ABS / MIN / MAX），零外部组件依赖
  同拍双窗配比  : tSwitchOverlap（重叠期）与 tSwitchInterval（轮值周期）同源于切换节奏；
                  配比约束 tSwitchOverlap < tSwitchInterval（组态闸强制），保证重叠期不会越过下一次轮值点

  码表 Error codes（本件格 03_2_0D，子码步进 +0x10）:
    16#0003_020D 故障级：组态非法（穿透门限 <= 0 / 轮值周期 <= 0 / 重叠期 <= 0 / 重叠期 >= 轮值周期）
    16#0003_021D 故障级：双塔均不可用（bBothFault 锁存）
    16#0003_022D 故障级：切换重叠期两塔同时离线（严重故障，独立归因）
    16#0003_023D 故障级：状态机落 ELSE 兜底（非法相位 ID）
    16#0003_010D 信息级：穿透超限提前切换（不置 bError）
    16#0003_011D 信息级：目标塔不可用，禁止切换并保持运行塔（不置 bError）
    16#0003_012D 信息级：轮值到点正常切换（不置 bError）
    16#0003_013D 信息级：压差反馈非有限，本拍不参与切换判据（不置 bError）

  修订历史 Revision :
    2026-11-18  v1.0.0  R37 首版
*)

TYPE E_DL_PurgeDutyState :
(
    eIdle      := 0,   // 空闲：未使能，双塔全停 / Idle, both towers off
    eRunA      := 10,  // A 塔值班 / Tower A online
    eRunB      := 20,  // B 塔值班 / Tower B online
    eSwitching := 30,  // 切换重叠：两塔同时在线（按允许处理）/ Switching overlap, both towers online
    eFault     := 90   // 故障：锁存待复位 / Fault, latched until reset
);
END_TYPE

FUNCTION_BLOCK FB_DL_VentPurgeDuty
VAR_INPUT
    bEnable         : BOOL := FALSE;           // 总使能，FALSE 时双塔全停 / Master enable, both towers off when low
    bReset          : BOOL := FALSE;           // 复位，上升沿清故障锁存 / Reset, rising edge clears the latch
    bTowerAAvail    : BOOL := FALSE;           // A 塔可用（无故障且再生完成）/ Tower A available
    bTowerBAvail    : BOOL := FALSE;           // B 塔可用（无故障且再生完成）/ Tower B available
    fTowerADpKpa    : REAL := 0.0;             // A 塔吸附压差 [kPa]，域 >= 0 / Tower A adsorption differential [kPa]
    fTowerBDpKpa    : REAL := 0.0;             // B 塔吸附压差 [kPa]，域 >= 0 / Tower B adsorption differential [kPa]
    fBreakthroughKpa : REAL := 3.5;            // 穿透门限 [kPa]，域 > 0 / Breakthrough threshold [kPa]
    tSwitchInterval : TIME := T#8H;            // 轮值周期（**小时口径**组态，内部换算 ms 计时）[h] / Duty interval configured in hours
    tSwitchOverlap  : TIME := T#30S;           // 切换重叠期（两塔同时在线）[ms]，域 > 0 且 < 轮值周期 / Switch overlap [ms]
    bForceSwitch    : BOOL := FALSE;           // 手动强制切换（上升沿受理，维修用）/ Manual forced switch, rising edge
END_VAR
VAR_OUTPUT
    bTowerAOnline   : BOOL;                    // A 塔在线 / Tower A online
    bSwitchCmd      : BOOL;                    // 切换指令（脉冲语义：置位 1 个 PLC 周期）/ Switch command, asserted for one PLC scan
    bBreakthroughWarn : BOOL;                  // 穿透告警（值班塔压差越门限）/ Breakthrough warning on the online tower
    bBothFault      : BOOL;                    // 双塔均不可用（锁存）/ Both towers unavailable, latched
    nSwitchCount    : UINT;                    // 累计切换次数 [次]，饱和不回绕 / Switch count, saturated, never wrapped
    fRemainSec      : REAL;                    // 本轮值班剩余时间 [s] / Remaining duty time [s]
    bValid          : BOOL;                    // 判据可用标志 / Criteria usable
    bError          : BOOL;                    // 故障标志，派生自锁存 / Fault flag derived from the latch
    nErrId          : UDINT;                   // 事件码，0 = 无事件 / Event code, 0 = no event
    eStateOut       : E_DL_PurgeDutyState;     // 状态出口，段尾单点映射 / State outlet, mapped at the tail
END_VAR
VAR
    tonDuty      : TON;                        // 轮值计时，每拍无条件调用 / Duty timer, called unconditionally
    tonOverlap   : TON;                        // 重叠期计时，每拍无条件调用 / Overlap timer, called unconditionally
    tonHeart     : TON;                        // 周期心跳窗，自复位 / Periodic heartbeat window, self-resetting
    rtReset      : R_TRIG;                     // 复位上升沿 / Reset rising edge
    rtForce      : R_TRIG;                     // 强制切换上升沿 / Forced switch rising edge
    _eState      : E_DL_PurgeDutyState := E_DL_PurgeDutyState.eIdle;  // 内部相位（CASE 唯一写入目标）/ Internal phase
    _uFault      : UDINT;                      // 故障码锁存 / Latched fault code
    _uInfo       : UDINT;                      // 信息码，每拍重算 / Information code, recomputed per scan
    _bFault      : BOOL;                       // 故障锁存位 / Latched fault bit
    _bBothFault  : BOOL;                       // 双塔不可用保持量 / Held both-unavailable value
    _bParamBad   : BOOL;                       // 组态非法聚合 / Configuration invalid aggregate
    _bAOnline    : BOOL;                       // A 塔在线内部量 / Internal tower A online
    _bBOnline    : BOOL;                       // B 塔在线内部量 / Internal tower B online
    _bToTowerA   : BOOL;                       // 切换目标塔（TRUE = 切往 A）/ Switch target, TRUE means tower A
    _bSwitchPulse: BOOL;                       // 内部切换单拍标志 → 段 8 映射 / Internal one-shot switch flag
    _bDpValidA   : BOOL;                       // A 塔压差有效 / Tower A differential usable
    _bDpValidB   : BOOL;                       // B 塔压差有效 / Tower B differential usable
    _bBreachA    : BOOL;                       // A 塔穿透 / Tower A broke through
    _bBreachB    : BOOL;                       // B 塔穿透 / Tower B broke through
    _bSwitchNeed : BOOL;                       // 本拍需要切换（到点 / 穿透 / 强制）/ A switch is due this scan
    _bOverlapBad : BOOL;                       // 重叠期两塔同时离线 / Both towers offline during the overlap
    _nCountAcc   : UINT;                       // 切换计数保持量 [次] / Held switch count
    _tIntervalMs : DINT;                       // 轮值周期毫秒值 [ms]，已钳位 / Duty interval in milliseconds, clamped
    _tOverlapMs  : DINT;                       // 重叠期毫秒值 [ms]，已钳位 / Overlap in milliseconds, clamped
    _bSwEntry    : BOOL;                       // 进入切换相首拍标志（单拍脉冲两段式）/ First-scan-in-switching flag
    _bHeartBrk   : BOOL := TRUE;               // 心跳窗断输入一拍 / One-scan heartbeat break
    _bDutyBrk    : BOOL := TRUE;               // 轮值计时断输入一拍（换塔重启）/ One-scan duty break to restart the timer
    _bOverlapBrk : BOOL := TRUE;               // 重叠计时断输入一拍 / One-scan overlap break
END_VAR
VAR CONSTANT
    DL_CNT_MAX_UINT : UINT := 65534;   // 切换计数饱和上限 [次]（留 1 防回绕）/ Saturation ceiling, one below the wrap
    DL_DP_LIM_KPA   : REAL := 1000.0;  // 压差有限性上限 [kPa] / Differential magnitude ceiling [kPa]
    DL_HEART_WINDOW : TIME := T#2S;    // 心跳观察窗 [ms]，自复位节拍 / Heartbeat window, self-resetting
    DL_INTERVAL_MAX_MS : DINT := 2147483000;  // 轮值周期毫秒上限（防 TIME 溢出）[ms] / Interval ceiling to avoid TIME overflow
    DL_EPS          : REAL := 1.0E-6;  // 判零容差 [1] / Zero tolerance
END_VAR

(* —— 段 0：定时器与边缘检测无条件周期刷新（R182：调用语句不得置于 IF / CASE 内） —— *)
rtReset(CLK := bReset);                                          // 复位上升沿，每拍必调
rtForce(CLK := bForceSwitch);                                    // 强制切换上升沿，每拍必调
tonHeart(IN := (NOT tonHeart.Q) AND (NOT _bHeartBrk), PT := DL_HEART_WINDOW);  // 心跳窗自复位
_bHeartBrk := FALSE;                                             // 断输入拍在调用后自清
tonDuty(IN := (((_eState = E_DL_PurgeDutyState.eRunA) OR (_eState = E_DL_PurgeDutyState.eRunB))
               AND (NOT _bDutyBrk)),
        PT := DINT_TO_TIME(_tIntervalMs));                       // 轮值计时（h 口径已换算为 ms）
_bDutyBrk := FALSE;                                              // 断输入拍在调用后自清（换塔时置位重启）
tonOverlap(IN := (_eState = E_DL_PurgeDutyState.eSwitching) AND (NOT _bOverlapBrk),
           PT := DINT_TO_TIME(_tOverlapMs));                     // 重叠期计时（表达式入参）
_bOverlapBrk := FALSE;                                           // 断输入拍在调用后自清

(* —— 段 1：单拍量预清零（计数 / 保持量 / 锁存不入清单，R187①） —— *)
_uInfo       := 16#0000_0000;   // 信息码每拍重算
bError       := FALSE;          // 故障出口每拍重算，段 7 由锁存派生
bValid       := FALSE;          // 可用标志缺省 FALSE
bSwitchCmd   := FALSE;          // 切换出口缺省 FALSE（脉冲宽度 = 1 拍）
bBreakthroughWarn := FALSE;     // 穿透告警缺省 FALSE
_bSwitchPulse := FALSE;         // 内部切换单拍标志预清零
_bParamBad   := FALSE;          // 组态非法预清零
_bSwitchNeed := FALSE;          // 切换需求预清零
_bOverlapBad := FALSE;          // 重叠离线标志预清零
_bDpValidA   := FALSE;          // A 塔压差有效标志预清零
_bDpValidB   := FALSE;          // B 塔压差有效标志预清零

(* —— 段 2：复位沿清锁存 + 按码专清（bBothFault 解除式见边界 ③） —— *)
IF rtReset.Q THEN
    IF bTowerAAvail OR bTowerBAvail THEN
        _bBothFault := FALSE;          // 解除式：复位 AND 至少一塔可用
    END_IF
    IF NOT _bBothFault THEN
        _bFault := FALSE;              // 双塔故障保持量已释放才清故障位
        _uFault := 16#0000_0000;       // 清锁存码
    END_IF
END_IF
IF (_uFault = 16#0003_021D) AND (NOT _bBothFault) THEN
    _uFault := 16#0000_0000;           // 按码专清：双塔不可用保持量已释放 → 对应码清除
    _bFault := FALSE;                  // 锁存位同步清
END_IF

(* —— 段 3：组态域闸（含 h 口径换算与上限钳位，覆盖全部换算引脚，R151） —— *)
_tIntervalMs := TIME_TO_DINT(tSwitchInterval);          // 轮值周期：TIME 以小时口径组态，转换即 ms [ms]
_tOverlapMs  := TIME_TO_DINT(tSwitchOverlap);           // 重叠期毫秒值 [ms]
IF (fBreakthroughKpa <> fBreakthroughKpa) OR (fBreakthroughKpa <= 0.0) THEN
    _bParamBad := TRUE;                                 // 穿透门限非法（切换判据的分母语义）
END_IF
IF _tIntervalMs <= 0 THEN
    _bParamBad := TRUE;                                 // 轮值周期 <= 0
END_IF
IF _tIntervalMs > DL_INTERVAL_MAX_MS THEN
    _tIntervalMs := DL_INTERVAL_MAX_MS;                 // 上限钳位（防 TIME 表示溢出）
END_IF
IF _tOverlapMs <= 0 THEN
    _bParamBad := TRUE;                                 // 重叠期 <= 0（两塔无交叠会瞬时断气）
END_IF
IF (_tIntervalMs > 0) AND (_tOverlapMs >= _tIntervalMs) THEN
    _bParamBad := TRUE;                                 // 重叠期 >= 轮值周期：重叠尚未结束就该再切（不可能组态）
END_IF
IF _bParamBad THEN
    _uFault := 16#0003_020D;                            // 故障级：组态非法
    _bFault := TRUE;                                    // 锁存位置位（复位沿可清）
    bError  := TRUE;                                    // 故障标志置位（R45 配对）
    _eState := E_DL_PurgeDutyState.eFault;              // 进故障相
END_IF

(* —— 段 4：压差有效性、穿透判据与切换需求 —— *)
_bDpValidA := (fTowerADpKpa = fTowerADpKpa) AND (fTowerADpKpa >= 0.0) AND (fTowerADpKpa <= DL_DP_LIM_KPA);  // A 塔压差有效
_bDpValidB := (fTowerBDpKpa = fTowerBDpKpa) AND (fTowerBDpKpa >= 0.0) AND (fTowerBDpKpa <= DL_DP_LIM_KPA);  // B 塔压差有效
IF (NOT _bDpValidA) OR (NOT _bDpValidB) THEN
    _uInfo := 16#0003_013D;                             // 信息级：压差非有限，本拍不参与切换判据
END_IF
_bBreachA := _bDpValidA AND (fTowerADpKpa > fBreakthroughKpa);  // A 塔穿透（仅有效值参与）
_bBreachB := _bDpValidB AND (fTowerBDpKpa > fBreakthroughKpa);  // B 塔穿透（仅有效值参与）
IF (_eState = E_DL_PurgeDutyState.eRunA) THEN
    bBreakthroughWarn := _bBreachA;                     // 在线塔为 A：告警跟随 A
ELSIF (_eState = E_DL_PurgeDutyState.eRunB) THEN
    bBreakthroughWarn := _bBreachB;                     // 在线塔为 B：告警跟随 B
END_IF

_bSwitchNeed := tonDuty.Q OR rtForce.Q OR
                ((_eState = E_DL_PurgeDutyState.eRunA) AND _bBreachA) OR
                ((_eState = E_DL_PurgeDutyState.eRunB) AND _bBreachB);  // 到点 / 强制 / 在线塔穿透
IF _bSwitchNeed AND tonDuty.Q THEN
    _uInfo := 16#0003_012D;                             // 信息级：轮值到点切换
ELSIF _bSwitchNeed AND (((_eState = E_DL_PurgeDutyState.eRunA) AND _bBreachA) OR
                        ((_eState = E_DL_PurgeDutyState.eRunB) AND _bBreachB)) THEN
    _uInfo := 16#0003_010D;                             // 信息级：穿透超限提前切换
END_IF

(* —— 段 5：双塔可用性归因（三岔：均可用 / 单塔可用 / 均不可用） —— *)
IF (NOT bTowerAAvail) AND (NOT bTowerBAvail) THEN
    _bBothFault := TRUE;                                // 双塔均不可用：保持量置位
    _uFault := 16#0003_021D;                            // 故障级：双塔均不可用
    _bFault := TRUE;                                    // 锁存
    bError  := TRUE;                                    // 故障标志置位（R45 配对）
    _eState := E_DL_PurgeDutyState.eFault;              // 进故障相
END_IF

(* —— 段 6：相位机（只做迁移与在线/切换单拍标志；出口在段 8） —— *)
CASE _eState OF

E_DL_PurgeDutyState.eIdle:
    _bAOnline := FALSE;                                 // 空闲：两塔全停（唯一清零点在本相）
    _bBOnline := FALSE;
    IF bEnable AND (NOT _bFault) AND (NOT _bParamBad) THEN
        IF bTowerAAvail THEN
            _eState := E_DL_PurgeDutyState.eRunA;       // 首轮启动：优先 A 塔
            _bAOnline := TRUE;                          // A 塔上线
            _bDutyBrk := TRUE;                          // 轮值计时从零开始
        ELSIF bTowerBAvail THEN
            _eState := E_DL_PurgeDutyState.eRunB;       // A 不可用：B 塔上线
            _bBOnline := TRUE;                          // B 塔上线
            _bDutyBrk := TRUE;                          // 轮值计时从零开始
        END_IF
    END_IF

E_DL_PurgeDutyState.eRunA:
    _bAOnline := TRUE;                                  // A 塔在线
    _bBOnline := FALSE;                                 // B 塔离线（非重叠期）
    IF (NOT bEnable) OR (NOT bTowerAAvail) THEN
        IF bTowerBAvail THEN
            _bToTowerA := FALSE;                        // A 失效：切往 B
            _eState := E_DL_PurgeDutyState.eSwitching;  // 进切换重叠
            _bSwEntry := TRUE;                          // 切换首拍标志置位（单拍脉冲）
            _bOverlapBrk := TRUE;                       // 重叠计时从零
        ELSE
            _uInfo := 16#0003_011D;                     // 信息级：目标塔不可用，禁止切换
            _eState := E_DL_PurgeDutyState.eIdle;       // 回空闲（无可用塔，段 5 已置 021D）
            _bAOnline := FALSE;
        END_IF
    ELSIF _bSwitchNeed THEN
        IF bTowerBAvail THEN
            _bToTowerA := FALSE;                        // 切往 B
            _eState := E_DL_PurgeDutyState.eSwitching;  // 进切换重叠
            _bSwEntry := TRUE;                          // 切换首拍标志置位（单拍脉冲）
            _bOverlapBrk := TRUE;                       // 重叠计时从零
        ELSE
            _uInfo := 16#0003_011D;                     // 信息级：B 不可用，保持 A 继续值班
            _bDutyBrk := TRUE;                          // 轮值计时重启（避免每拍重复判到点）
        END_IF
    END_IF

E_DL_PurgeDutyState.eRunB:
    _bAOnline := FALSE;                                 // A 塔离线（非重叠期）
    _bBOnline := TRUE;                                  // B 塔在线
    IF (NOT bEnable) OR (NOT bTowerBAvail) THEN
        IF bTowerAAvail THEN
            _bToTowerA := TRUE;                         // B 失效：切往 A
            _eState := E_DL_PurgeDutyState.eSwitching;  // 进切换重叠
            _bSwEntry := TRUE;                          // 切换首拍标志置位（单拍脉冲）
            _bOverlapBrk := TRUE;                       // 重叠计时从零
        ELSE
            _uInfo := 16#0003_011D;                     // 信息级：目标塔不可用，禁止切换
            _eState := E_DL_PurgeDutyState.eIdle;       // 回空闲
            _bBOnline := FALSE;
        END_IF
    ELSIF _bSwitchNeed THEN
        IF bTowerAAvail THEN
            _bToTowerA := TRUE;                         // 切往 A
            _eState := E_DL_PurgeDutyState.eSwitching;  // 进切换重叠
            _bSwEntry := TRUE;                          // 切换首拍标志置位（单拍脉冲）
            _bOverlapBrk := TRUE;                       // 重叠计时从零
        ELSE
            _uInfo := 16#0003_011D;                     // 信息级：A 不可用，保持 B 继续值班
            _bDutyBrk := TRUE;                          // 轮值计时重启
        END_IF
    END_IF

E_DL_PurgeDutyState.eSwitching:
    _bAOnline := TRUE;                                  // 重叠期：两塔同时在线（按允许处理）
    _bBOnline := TRUE;
    IF _bSwEntry THEN
        _bSwitchPulse := TRUE;                          // 切换指令单拍：仅进入本相首拍置位，次拍段 1 清
        _bSwEntry := FALSE;                             // 首拍标志自清（唯一置假点）
    END_IF
    IF (NOT bTowerAAvail) AND (NOT bTowerBAvail) THEN
        _bOverlapBad := TRUE;                           // 重叠期两塔均不可用：严重故障（独立归因）
        _uFault := 16#0003_022D;                        // 故障级：重叠期两塔同时离线
        _bFault := TRUE;                                // 锁存
        bError  := TRUE;                                // 故障标志置位（R45 配对）
        _bAOnline := FALSE;                             // 安全侧：两塔全停
        _bBOnline := FALSE;
        _eState := E_DL_PurgeDutyState.eFault;          // 进故障相
    ELSIF tonOverlap.Q THEN
        _bAOnline := _bToTowerA;                        // 重叠结束：仅目标塔保持在线
        _bBOnline := NOT _bToTowerA;
        IF _nCountAcc < DL_CNT_MAX_UINT THEN
            _nCountAcc := _nCountAcc + 1;               // 切换计数 +1（饱和不回绕）
        END_IF
        IF _bToTowerA THEN
            _eState := E_DL_PurgeDutyState.eRunA;       // 目标 A：进 A 值班相
        ELSE
            _eState := E_DL_PurgeDutyState.eRunB;       // 目标 B：进 B 值班相
        END_IF
        _bDutyBrk := TRUE;                              // 新一轮轮值计时从零
    END_IF

E_DL_PurgeDutyState.eFault:
    _bAOnline := FALSE;                                 // 故障：两塔全停（安全侧）
    _bBOnline := FALSE;
    IF (NOT _bFault) AND (NOT _bParamBad) AND bEnable THEN
        _eState := E_DL_PurgeDutyState.eIdle;           // 锁存已清且组态合法：回空闲重新选塔
    END_IF

ELSE
    _uFault := 16#0003_023D;                            // 故障级：相位 ID 越界（枚举兜底）
    _bFault := TRUE;                                    // 锁存
    bError  := TRUE;                                    // 故障标志置位（R45 配对）
    _bAOnline := FALSE;                                 // 兜底安全侧：两塔全停
    _bBOnline := FALSE;
    _eState := E_DL_PurgeDutyState.eFault;              // 强制回故障相
END_CASE

(* —— 段 7：故障码优先级链与在线镜像仲裁（每个 bError 置位源在此均有码，R45） —— *)
IF _bParamBad THEN
    bError := TRUE;                                     // 组态非法：码已在段 3 置位（020D）
END_IF
IF _bOverlapBad AND (NOT _bFault) THEN
    _uFault := 16#0003_022D;                            // 独立归因：重叠期离线（即使其它码未置）
    _bFault := TRUE;                                    // 锁存
    bError  := TRUE;                                    // 故障标志置位（R45 配对）
    _bAOnline := FALSE;                                 // 安全侧
    _bBOnline := FALSE;
END_IF

(* —— 段 8：出口单点映射（名实同源；锁存码回放，禁同拍抹除） —— *)
bTowerAOnline := _bAOnline;                             // A 塔在线出口
bSwitchCmd    := _bSwitchPulse;                         // 切换指令出口：宽度恰 1 个 PLC 周期
bBothFault    := _bBothFault;                           // 双塔不可用出口（保持量）
nSwitchCount  := _nCountAcc;                            // 切换计数出口（UINT，饱和）
IF _tIntervalMs > 0 THEN
    fRemainSec := (DINT_TO_REAL(_tIntervalMs) - TIME_TO_REAL(tonDuty.ET)) / 1000.0;  // 剩余秒数（分母已证 > 0）
ELSE
    fRemainSec := 0.0;                                  // 组态非法：剩余时间无意义，置 0
END_IF
IF fRemainSec < 0.0 THEN
    fRemainSec := 0.0;                                  // 下限保护（到点后不出现负剩余）
END_IF
eStateOut := _eState;                                   // 状态出口
IF _bFault THEN
    nErrId := _uFault;                                  // 故障锁存码回放（不在故障相按当下输入重推）
    bError := TRUE;                                     // 故障出口派生自锁存
ELSE
    nErrId := _uInfo;                                   // 信息码
END_IF
bValid := bEnable AND (NOT _bFault) AND (NOT _bParamBad);  // 判据可用

END_FUNCTION_BLOCK
